RoboDK station: Celda_Soldadura_Estator_Grupo4_v05.rdk

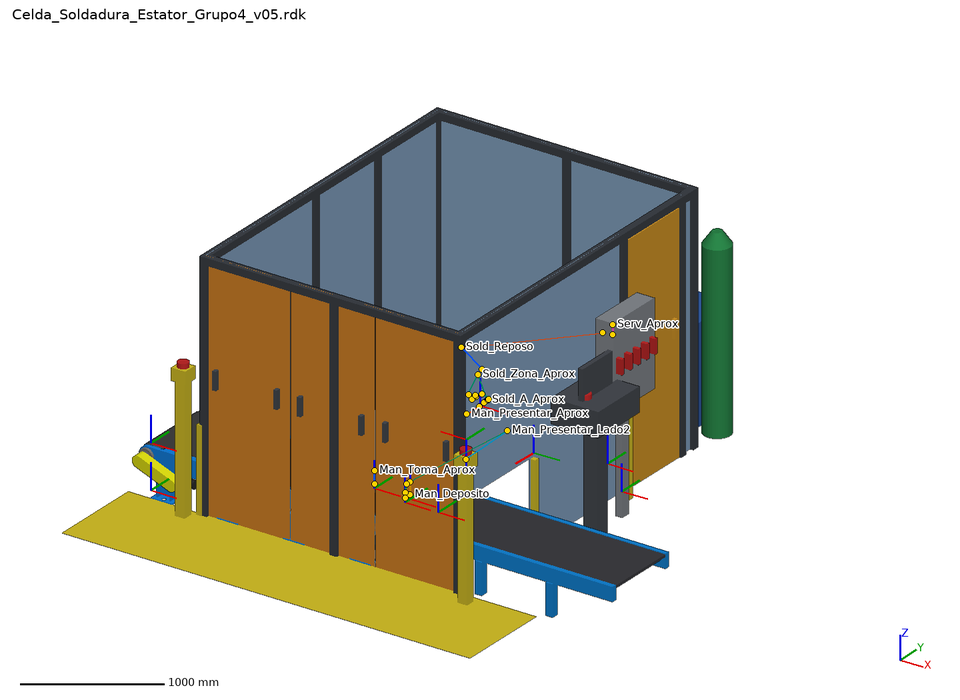
[picture v0: the station drawn from its stored meshes, robots at their saved joint values, targets as dots, program paths as lines]
Station Celda_Soldadura_Estator_Grupo4_v05 (saved by RoboDK 6.1.1). Poses are relative to the parent item; angles as X-Y-Z fixed-axis rotations.
Station parameters (name, value as stored): PIEZA_EN_TOMA, 0, PIEZA_PRESENTADA, 0, ARCO_TIG, 0, SOLDADURA_TERMINADA, 0, COORDINADOR_ACTIVO, 1, PERMISO_OPERACION, 0, ARRANQUE_ID, 0, ARRANQUE_ACK, 0, PARADA_ID, 0, PARADA_ACK, 0, AUTO_ACTIVO, 0, ESTADO_CONTROL, 0, CAUSA_RECHAZO, 0, PROXIMA_PIEZA, 1, PIEZA_ACTIVA, 0, CELDA_INICIALIZADA, 0, PIEZAS_COMPLETADAS, 0, LOTES_COMPLETADOS, 0, MODO_ID, 0, MODO_ACK, 0, MODO_SOLICITADO, 0, MODO_CONFIRMADO, 0, MODO_OBJETIVO, 0, MODO_EN_TRANSICION, 0, MODO_RESULTADO, 0, MODO_CAUSA, 0, MODO_ID_CAPTURADO, 0, MODO_CAPTURADO, 0, MODO_DESDE_AUTO, 0, MODO_ES_INTERVENCION, 0, MODO_CONOCIDO, 0, SENSORES_VALIDOS, 0, PIEZA_SUJETA_SENSOR, 0, IRB_EN_REPOSO, 0, CRB_EN_REPOSO, 0, IRB_EN_MANT, 0, CRB_EN_MANT, 0, CRB_EN_SERVICIO, 0, CINTA_DETENIDA, 0, IRB_DISPONIBLE, 0, CRB_DISPONIBLE, 0, CINTA_DISPONIBLE, 0, CONF_RESTITUCION, 0, FASE_PIEZA, 0, FASE_CAPTURADA, 0, PARO_CAUSA, 0, RECUP_PENDIENTE, 0, RECUPERAR_ID, 0, RECUPERAR_ACK, 0, PIEZAS_RETRABAJO, 0, RETRABAJO_ACTUAL, 0, SUJETA_CAPTURADA, 0, PIEZA_RESUELTA, 0, EMERGENCIA_SIM, 0, CORTINA_ENTRADA_SIM, 0, CORTINA_SALIDA_SIM, 0, PUERTA_ABIERTA_SIM, 0, OBJETIVO_PIEZAS, 0, PIEZAS_BUENAS, 0, PEDIDO_CUMPLIDO, 0, PEDIDOS_TERMINADOS, 0, REINICIAR_ID, 0, REINICIAR_ACK, 0, PEDIDO_PARADA, 0
  - frame Frame_Celda at (0, 0, 0) mm
    - frame Base_Manipulador_IRB1200 at (0, 0, 0) mm
      - robot ABB IRB 1200-7/0.7: 6 axes, payload 7 kg, reach 703 mm, repeatability 0.02 mm, weight 54 kg
          modified DH rows (alpha deg, a mm, theta deg, d mm): 0, 0, 0, 399; -90, 0, -90, 0; 0, 350, 0, 0; -90, 42, 0, 351; 90, 0, 0, 0; -90, 0, 180, 82
          joint limits [-170, -100, -200, -270, -130, -360] to [170, 135, 70, 270, 130, 360]; home [0, 0, 0, 0, 0, 0]; saved at [0, -20, 30, 0, 80, 0]
        - frame RobotiQ 2F-85 Gripper (Mechanism) Base at (0, 0, 0) mm
          - robot Pinza_2F85 (model RobotiQ 2F85): 1 axes, payload 5 kg
              joint limits [0] to [85]; home [85]; saved at [85]
        - tool TCP_Pinza, TCP at (0, 0, 150) mm
    - frame Base_Soldador_CRB1300 at (0, 1150, 0) mm, rotated rx 0 ry 0 rz -90 deg
      - robot ABB CRB 1300-10/1.15: 6 axes
          modified DH rows (alpha deg, a mm, theta deg, d mm): 0, 0, 0, 544; -90, 150, -90, 0; 0, 575, 0, 0; -90, 40, 0, 425; 90, 0, 0, 0; -90, 0, 180, 90
          joint limits [-180, -95, -210, -230, -130, -242] to [180, 155, 65, 230, 130, 242]; home [0, 0, 0, 0, 0, 0]; saved at [0, -10, 10, 0, 60, 0]
        - tool Antorcha_TIG, TCP at (0, 0, 207) mm, size 80 x 80 x 207 mm, geometry from antorcha_tig.stl
    - frame Base_Cinta_Pasante at (-1830, -860, 0) mm
      - robot Cinta_Pasante: 1 axes
          modified DH rows (alpha deg, a mm, theta deg, d mm): 0, 0, 0, 0 linear
          base shift (0, 0, 0) mm, rotated rx 0 ry 90 rz 0 deg
          joint limits [-900000] to [900000]; home [0]; saved at [0]
        - frame Frame_Banda at (0, 0, 0) mm
          - frame Frame_Piezas_Soldadas at (0, 0, 0) mm
          - object Estator_1 at (1680, 300, 0) mm, size 105 x 105 x 55 mm, geometry from paquete_estator.stl
          - object Estator_2 at (1380, 300, 0) mm, size 105 x 105 x 55 mm, geometry from paquete_estator.stl
          - object Estator_3 at (1080, 300, 0) mm, size 105 x 105 x 55 mm, geometry from paquete_estator.stl
          - object Estator_4 at (780, 300, 0) mm, size 105 x 105 x 55 mm, geometry from paquete_estator.stl
    - object Sensor_Pieza_En_Toma at (-150, -900, 396.5) mm, rotated rx 0 ry 0 rz 90 deg, size 683.3 x 45.2 x 12.5 mm, geometry from Laser-Sensor.stl
    - object Estacion_Servicio_Antorcha at (520, 1300, 0) mm, size 250 x 250 x 1000 mm, geometry from estacion_servicio_antorcha.stl
    - frame Frame_Cerramiento at (0, 0, 0) mm
      - frame Bisagra_Puerta at (850, 1000, 0) mm
        - object Puerta at (0, 0, 0) mm, size 60 x 700 x 1920 mm, geometry from puerta.stl
      - object Cerramiento_Estructura at (0, 0, 0) mm, size 2210 x 2870 x 2000 mm, geometry from cerramiento_estructura_v04.stl
      - object Cerramiento_Paneles at (0, 0, 0) mm, size 2154 x 2812 x 2000 mm, geometry from cerramiento_paneles_v04.stl
      - object Paneles_Desmontables_Sur at (0, 0, 0) mm, size 2140 x 4 x 2000 mm, geometry from paneles_desmontables_sur.stl
      - object Paneles_Desmontables_Manijas at (0, 0, 0) mm, size 1980 x 38 x 150 mm, geometry from paneles_desmontables_manijas.stl
      - object Cortina_Luz_Entrada at (-1330, 0, 0) mm, size 40 x 920 x 700 mm, geometry from cortina_luz_cinta_v04.stl
      - object Cortina_Luz_Salida at (880, 0, 0) mm, size 40 x 920 x 700 mm, geometry from cortina_luz_cinta_v04.stl
    - frame Frame_Soldadura at (0, 500, 620) mm
      - target Man_Presentar_Aprox (joint target) at (0, -157.5, 0) mm, rotated rx -90 ry 0 rz 0 deg; joints [90, -43.636, 55.703, 0, -12.068, -90] of ABB IRB 1200-7/0.7
      - target Man_Presentar_Lado1 (joint target) at (0, -7.5, 0) mm, rotated rx -90 ry 0 rz 0 deg; joints [90, -11.774, 38.724, 0, -26.95, -90] of ABB IRB 1200-7/0.7
      - target Man_Presentar_Lado2 (joint target) at (583, -500, 171) mm, rotated rx 0 ry 90 rz 0 deg; joints [90, -11.774, 38.724, 0, -26.95, 90] of ABB IRB 1200-7/0.7
      - target Man_Presentar_Aprox_Lado2 (joint target) at (583, -500, 171) mm, rotated rx 0 ry 90 rz 0 deg; joints [90, -43.636, 55.703, 0, -12.068, 90] of ABB IRB 1200-7/0.7
      - target Sold_Zona_Aprox (Cartesian target) at (0, -26.5, 250) mm, rotated rx 180 ry 0 rz 90 deg; joints [103.36, 41.617, 53.414, 0, -5.031, 103.36] of ABB CRB 1300-10/1.15
      - target Sold_A_Aprox (Cartesian target) at (78.2, -26.5, 78.2) mm, rotated rx -135 ry 0 rz 90 deg; joints [98.688, 74.302, 5.58, 7.491, 55.018, 91.856] of ABB CRB 1300-10/1.15
      - target Sold_A_Inicio (Cartesian target) at (49.91, -26.5, 49.91) mm, rotated rx -135 ry 0 rz 90 deg; joints [98.998, 76.411, 8.063, 8.245, 50.464, 91.119] of ABB CRB 1300-10/1.15
      - target Sold_A_Fin (Cartesian target) at (49.91, 26.5, 49.91) mm, rotated rx -135 ry 0 rz 90 deg; joints [102.751, 76.611, 6.557, 11.474, 51.681, 91.918] of ABB CRB 1300-10/1.15
      - target Sold_Transicion_Medio (Cartesian target) at (0, 26.5, 80) mm, rotated rx 180 ry 0 rz 90 deg; joints [108.748, 65.119, 46.933, 0, -22.052, 108.748] of ABB CRB 1300-10/1.15
      - target Sold_B_Inicio (Cartesian target) at (-49.91, 26.5, 49.91) mm, rotated rx 135 ry 0 rz 90 deg; joints [124.163, 102.688, 60.997, 205.222, 111.278, -54.665] of ABB CRB 1300-10/1.15
      - target Sold_B_Fin (Cartesian target) at (-49.91, -26.5, 49.91) mm, rotated rx 135 ry 0 rz 90 deg; joints [115.401, 107.202, 62.682, 200.569, 120.307, -60.716] of ABB CRB 1300-10/1.15
      - target Sold_B_Retiro (Cartesian target) at (-78.2, -26.5, 78.2) mm, rotated rx 135 ry 0 rz 90 deg; joints [-61.951, -75.264, -208.995, 23.114, 57.885, -82.141] of ABB CRB 1300-10/1.15
      - target Sold_A_Salida (Cartesian target) at (56.57, 26.5, 56.57) mm, rotated rx -135 ry 0 rz 90 deg; joints [102.647, 76.107, 6.003, 11.22, 52.72, 92.165] of ABB CRB 1300-10/1.15
      - target Sold_B_Entrada (Cartesian target) at (-56.57, 26.5, 56.57) mm, rotated rx 135 ry 0 rz 90 deg; joints [124.856, 103.181, 62.152, 205.935, 112.476, -53.248] of ABB CRB 1300-10/1.15
    - frame Frame_Toma_Cinta at (-150, -560, 366.5) mm
      - target Man_Toma_Aprox (joint target) at (0, 0, 135) mm, rotated rx 180 ry 0 rz 0 deg; joints [-104.995, 41.989, -47.307, 0, 95.319, 75.005] of ABB IRB 1200-7/0.7
      - target Man_Toma (joint target) at (0, 0, 35) mm, rotated rx 180 ry 0 rz 0 deg; joints [-104.995, 40.57, -28.656, 0, 78.086, 75.005] of ABB IRB 1200-7/0.7
    - frame Frame_Servicio at (520, 1300, 0) mm
      - target Serv_Aprox (Cartesian target) at (0, 60, 1050) mm, rotated rx 180 ry 0 rz 0 deg; joints [-125.65, 36.775, -52.607, 69.175, 38.577, -64.055] of ABB CRB 1300-10/1.15
      - target Serv_Verificacion_TCP (Cartesian target) at (0, 60, 973) mm, rotated rx 180 ry 0 rz 0 deg; joints [-125.65, 36.775, -52.607, 69.175, 38.577, -64.055] of ABB CRB 1300-10/1.15
      - target Serv_Cambio_Tungsteno (Cartesian target) at (0, -65, 1035) mm, rotated rx 180 ry 0 rz 0 deg; joints [-125.65, 36.775, -52.607, 69.175, 38.577, -64.055] of ABB CRB 1300-10/1.15
    - target Man_Reposo (joint target) at (583, 0, 791) mm, rotated rx 0 ry 90 rz 0 deg; joints [0, -20, 30, 0, 80, 0] of ABB IRB 1200-7/0.7
    - target Sold_Reposo (joint target) at (0, 278, 1159) mm, rotated rx 0 ry 90 rz -90 deg; joints [0, -10, 10, 0, 60, 0] of ABB CRB 1300-10/1.15
    - target Pinza_Abierta (joint target) at (536.92, 0, 791) mm, rotated rx 0 ry 90 rz 0 deg; joints [85] of Pinza_2F85
    - target Pinza_Cerrada (joint target) at (536.92, 0, 791) mm, rotated rx 0 ry 90 rz 0 deg; joints [0] of Pinza_2F85
    - target Pinza_Sujeta (joint target) at (536.92, 0, 791) mm, rotated rx 0 ry 90 rz 0 deg; joints [35] of Pinza_2F85
    - target Cinta_Posicion_1 (joint target) at (-1830, -860, 366.5) mm; joints [0] of Cinta_Pasante
    - target Cinta_Posicion_2 (joint target) at (-1830, -860, 366.5) mm; joints [300] of Cinta_Pasante
    - target Cinta_Posicion_3 (joint target) at (-1830, -860, 366.5) mm; joints [600] of Cinta_Pasante
    - target Cinta_Posicion_4 (joint target) at (-1830, -860, 366.5) mm; joints [900] of Cinta_Pasante
    - object Cinta_Salida_Banda at (0, 0, 0) mm, size 1880 x 600 x 20 mm, geometry from cinta_extension_banda.stl
    - object Cinta_Salida_Estructura at (0, 0, 0) mm, size 1880 x 700 x 371.5 mm, geometry from cinta_extension_estructura.stl
    - frame Frame_Deposito_Cinta at (150, -560, 366.5) mm
      - target Man_Deposito_Aprox (Cartesian target) at (0, 0, 135) mm, rotated rx 180 ry 0 rz 0 deg; joints [0, -20, 30, 0, 80, 0] of ABB IRB 1200-7/0.7
      - target Man_Deposito (Cartesian target) at (0, 0, 35) mm, rotated rx 180 ry 0 rz 0 deg; joints [0, -20, 30, 0, 80, 0] of ABB IRB 1200-7/0.7
    - target Cinta_Evacuacion (joint target) at (-1830, -860, 366.5) mm; joints [1750] of Cinta_Pasante
    - object Pasillo_Mantenimiento at (0, 0, 0) mm, size 3450 x 800 x 3 mm, geometry from pasillo_mantenimiento.stl
    - object Accionamiento_Cinta at (-1760, -80, 0) mm, size 140 x 320 x 296.5 mm, geometry from accionamiento_cinta.stl
    - object Accionamiento_Cinta_Resguardo at (-1760, -80, 0) mm, size 220 x 400 x 200 mm, geometry from accionamiento_cinta_resguardo.stl
    - object Tablero_LOTO at (1010, 700, 0) mm, size 150 x 500 x 1600 mm, geometry from tablero_loto.stl
    - object Tablero_LOTO_Seccionadores at (1010, 700, 0) mm, size 50 x 430 x 120 mm, geometry from tablero_loto_manijas.stl
    - object Panel_Operador at (1150, 250, 0) mm, size 400 x 500 x 1400 mm, geometry from panel_operador.stl
    - object Parada_Emergencia_Panel at (1150, 130, 0) mm, size 90 x 90 x 40 mm, geometry from parada_emergencia_hongo.stl
    - object Parada_Emergencia_Puerta_Poste at (930, 920, 0) mm, size 120 x 120 x 1150 mm, geometry from parada_emergencia_poste.stl
    - object Parada_Emergencia_Puerta at (930, 920, 0) mm, size 90 x 90 x 40 mm, geometry from parada_emergencia_hongo.stl
    - object Parada_Emergencia_Entrada_Poste at (-1420, -1060, 0) mm, size 120 x 120 x 1150 mm, geometry from parada_emergencia_poste.stl
    - object Parada_Emergencia_Entrada at (-1420, -1060, 0) mm, size 90 x 90 x 40 mm, geometry from parada_emergencia_hongo.stl
    - object Parada_Emergencia_Salida_Poste at (970, -1060, 0) mm, size 120 x 120 x 1150 mm, geometry from parada_emergencia_poste.stl
    - object Parada_Emergencia_Salida at (970, -1060, 0) mm, size 90 x 90 x 40 mm, geometry from parada_emergencia_hongo.stl
    - object Controlador_IRB1200 at (-800, 1950, 0) mm, size 600 x 500 x 1200 mm, geometry from gabinete_controlador.stl
    - object Controlador_CRB1300 at (-100, 1950, 0) mm, size 600 x 500 x 1200 mm, geometry from gabinete_controlador.stl
    - object Fuente_TIG at (500, 1950, 0) mm, size 400 x 600 x 800 mm, geometry from fuente_tig.stl
    - object Cilindro_Argon at (850, 2150, 0) mm, size 220 x 220 x 1550 mm, geometry from cilindro_argon.stl
    - target Man_Mantenimiento (joint target) at (233.25, 0, 476.3) mm, rotated rx 180 ry 0 rz -180 deg; joints [45, -30, 50, 0, 60, 0] of ABB IRB 1200-7/0.7
    - target Sold_Mantenimiento (joint target) at (0, 526.35, 893.05) mm, rotated rx 180 ry 30 rz 90 deg; joints [100, -30, 50, 0, 60, 0] of ABB CRB 1300-10/1.15
    - frame Frame_Deposito_Retrabajo at (150, -620, 366.5) mm
      - target Man_Retrabajo_Aprox (Cartesian target) at (0, 20, 135) mm, rotated rx 180 ry 0 rz 0 deg; joints [14.425, -18.655, 29.096, 0, 79.558, 14.425] of ABB IRB 1200-7/0.7
      - target Man_Retrabajo_Salida (Cartesian target) at (0, 0, 75) mm, rotated rx 180 ry 0 rz 0 deg; joints [14.425, -18.655, 29.096, 0, 79.558, 14.425] of ABB IRB 1200-7/0.7
      - target Man_Retrabajo (Cartesian target) at (0, 0, 35) mm, rotated rx 180 ry 0 rz 0 deg; joints [14.425, -18.655, 29.096, 0, 79.558, 14.425] of ABB IRB 1200-7/0.7
  - program Pinza_Abrir (2 instructions, listed below)
  - program Pinza_Cerrar (2 instructions, listed below)
  - program Pinza_Sujetar (2 instructions, listed below)
  - program Cinta_Avanzar_1 (4 instructions, listed below)
  - program Cinta_Avanzar_2 (4 instructions, listed below)
  - program Cinta_Avanzar_3 (4 instructions, listed below)
  - program Cinta_Avanzar_4 (4 instructions, listed below)
  - program Evento_Tomar_Pieza (2 instructions, listed below)
  - program Evento_Soltar_Pieza (2 instructions, listed below)
  - program Man_Ir_Reposo (4 instructions, listed below)
  - program Man_Tomar_Cinta (16 instructions, listed below)
  - program Man_Presentar_Lado1 (8 instructions, listed below)
  - program Man_Presentar_Lado2 (8 instructions, listed below)
  - program Sold_Ir_Reposo (4 instructions, listed below)
  - program Sold_Par_Cordones (38 instructions, listed below)
  - program Sold_Servicio_Antorcha (10 instructions, listed below)
  - program Inicio_Celda (8 instructions, listed below)
  - program Ciclo_Pieza_1 (15 instructions, listed below)
  - program Ciclo_Pieza_2 (15 instructions, listed below)
  - program Ciclo_Pieza_3 (15 instructions, listed below)
  - program Ciclo_Pieza_4 (17 instructions, listed below)
  - program Fin_Lote (6 instructions, listed below)
  - program Programa_Principal (8 instructions, listed below)
  - program Man_Depositar_Cinta (18 instructions, listed below)
  - program Cinta_Evacuar (2 instructions, listed below)
  - program Man_Ir_Mantenimiento (7 instructions, listed below)
  - program Sold_Ir_Mantenimiento (7 instructions, listed below)
  - program Preparar_Servicio_Antorcha (5 instructions, listed below)
  - program Parada_Entre_Piezas (7 instructions, listed below)
  - program Atender_Solicitud_Modo (598 instructions, listed below)
  - program Confirmar_Posicion_Modo (113 instructions, listed below)
  - program Man_Depositar_Retrabajo (19 instructions, listed below)
  - program Sold_Retirar (5 instructions, listed below)
  - program Recuperar_Desde_Lado1 (21 instructions, listed below)
  - program Recuperar_Desde_Lado2 (20 instructions, listed below)
  - program Recuperar_Deposito (18 instructions, listed below)
  - program Recuperar_Pieza (97 instructions, listed below)
  - program Cerrar_Pedido (14 instructions, listed below)
  - program Coordinador_Panel (275 instructions, listed below)
  - Python program Abrir_Panel_Operador (listed below)
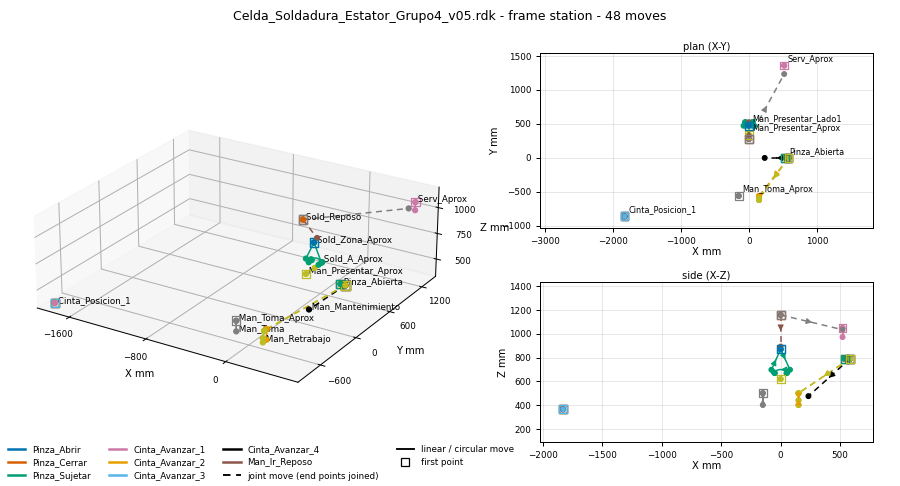
[picture p0: tool path of Celda_Soldadura_Estator_Grupo4_v05.rdk in frame station, 48 of 48 moves have a stored position in this frame; points joined in program order, loops and branches not executed]

--- program Pinza_Abrir (robot Pinza_2F85) ---
  Apertura máxima: reposo de la pinza
  MoveJ (Pinza_Abierta)

--- program Pinza_Cerrar (robot Pinza_2F85) ---
  Dedos juntos para entrar o salir del agujero del estator
  MoveJ (Pinza_Cerrada)

--- program Pinza_Sujetar (robot Pinza_2F85) ---
  Agarre interior: los dedos se abren contra el agujero de Ø55
  MoveJ (Pinza_Sujeta)

--- program Cinta_Avanzar_1 (robot Cinta_Pasante) ---
  Lleva el estator 1 del lote a la posición de toma
  MoveJ (Cinta_Posicion_1)
  Señal del sensor láser: hay pieza en la toma
  Set PIEZA_EN_TOMA=1

--- program Cinta_Avanzar_2 (robot Cinta_Pasante) ---
  Lleva el estator 2 del lote a la posición de toma
  MoveJ (Cinta_Posicion_2)
  Señal del sensor láser: hay pieza en la toma
  Set PIEZA_EN_TOMA=1

--- program Cinta_Avanzar_3 (robot Cinta_Pasante) ---
  Lleva el estator 3 del lote a la posición de toma
  MoveJ (Cinta_Posicion_3)
  Señal del sensor láser: hay pieza en la toma
  Set PIEZA_EN_TOMA=1

--- program Cinta_Avanzar_4 (robot Cinta_Pasante) ---
  Lleva el estator 4 del lote a la posición de toma
  MoveJ (Cinta_Posicion_4)
  Señal del sensor láser: hay pieza en la toma
  Set PIEZA_EN_TOMA=1

--- program Evento_Tomar_Pieza (robot ABB IRB 1200-7/0.7) ---
  Engancha a TCP_Pinza el estator que la pinza acaba de sujetar
  Adjuntar a TCP_Pinza

--- program Evento_Soltar_Pieza (robot ABB IRB 1200-7/0.7) ---
  Libera el estator sobre la banda (Frame_Piezas_Soldadas)
  Separar de TCP_Pinza

--- program Man_Ir_Reposo (robot ABB IRB 1200-7/0.7) ---
  Posición de reposo fuera de la zona de soldadura
  Est. herr: TCP_Pinza
  Establecer velocidad (1000.0 mm/s)
  MoveJ (Man_Reposo)

--- program Man_Tomar_Cinta (robot ABB IRB 1200-7/0.7) ---
  Toma el estator de la cinta con agarre interior
  Est. Ref.: Frame_Toma_Cinta
  Est. herr: TCP_Pinza
  Wait PIEZA_EN_TOMA=1
  Establecer velocidad (1000.0 mm/s)
  Suave(5)
  MoveJ (Man_Toma_Aprox)
  Llamar Pinza_Cerrar
  Suave(0)
  Establecer velocidad (100.0 mm/s)
  Entrada vertical en el agujero: MoveL para no rozar la pieza
  MoveL (Man_Toma)
  Llamar Pinza_Sujetar
  Llamar Evento_Tomar_Pieza
  Set PIEZA_EN_TOMA=0
  MoveL (Man_Toma_Aprox)

--- program Man_Presentar_Lado1 (robot ABB IRB 1200-7/0.7) ---
  Presenta las aristas A y B arriba, con el eje del estator hacia el soldador
  Est. Ref.: Frame_Soldadura
  Est. herr: TCP_Pinza
  Establecer velocidad (1000.0 mm/s)
  MoveJ (Man_Presentar_Aprox)
  Establecer velocidad (100.0 mm/s)
  MoveL (Man_Presentar_Lado1)
  Set PIEZA_PRESENTADA=1

--- program Man_Presentar_Lado2 (robot ABB IRB 1200-7/0.7) ---
  Gira 180° sobre el eje de la pinza (J6) para subir las aristas C y D
  Est. Ref.: Frame_Soldadura
  Est. herr: TCP_Pinza
  Wait SOLDADURA_TERMINADA=1
  Set SOLDADURA_TERMINADA=0
  Establecer velocidad (100.0 mm/s)
  MoveJ (Man_Presentar_Lado2)
  Set PIEZA_PRESENTADA=1

--- program Sold_Ir_Reposo (robot ABB CRB 1300-10/1.15) ---
  Reposo del soldador fuera del volumen de giro de la pieza
  Est. herr: Antorcha_TIG
  Establecer velocidad (1000.0 mm/s)
  MoveJ (Sold_Reposo)

--- program Sold_Par_Cordones (robot ABB CRB 1300-10/1.15) ---
  Suelda las dos aristas superiores del estator presentado
  Est. Ref.: Frame_Soldadura
  Est. herr: Antorcha_TIG
  Wait PIEZA_PRESENTADA=1
  Establecer velocidad (1000.0 mm/s)
  Suave(5)
  MoveJ (Sold_Zona_Aprox)
  Suave(0)
  Establecer velocidad (300.0 mm/s)
  Aproximación radial a la arista A
  MoveL (Sold_A_Aprox)
  Establecer velocidad (100.0 mm/s)
  MoveL (Sold_A_Inicio)
  Cordón A: arco encendido, avance recto a velocidad de soldadura
  Set ARCO_TIG=1
  Establecer velocidad (5.0 mm/s)
  MoveL (Sold_A_Fin)
  Set ARCO_TIG=0
  Establecer velocidad (100.0 mm/s)
  Separación radial: la punta sale del escalón antes de rodear la pieza
  MoveL (Sold_A_Salida)
  Establecer velocidad (200.0 mm/s)
  Transición en arco alrededor del eje del estator, a radio constante
  MoveC (Sold_Transicion_Medio, Sold_B_Entrada)
  Establecer velocidad (100.0 mm/s)
  MoveL (Sold_B_Inicio)
  Cordón B: avance recto en sentido contrario al A
  Set ARCO_TIG=1
  Establecer velocidad (5.0 mm/s)
  MoveL (Sold_B_Fin)
  Set ARCO_TIG=0
  Establecer velocidad (200.0 mm/s)
  MoveL (Sold_B_Retiro)
  Establecer velocidad (300.0 mm/s)
  MoveL (Sold_Zona_Aprox)
  Set PIEZA_PRESENTADA=0
  Set SOLDADURA_TERMINADA=1
  Llamar Sold_Ir_Reposo

--- program Sold_Servicio_Antorcha (robot ABB CRB 1300-10/1.15) ---
  Verificación del TCP al final de cada lote
  Est. Ref.: Frame_Servicio
  Est. herr: Antorcha_TIG
  Establecer velocidad (500.0 mm/s)
  MoveJ (Serv_Aprox)
  Establecer velocidad (100.0 mm/s)
  Bajada vertical hasta el cruce de los haces
  MoveL (Serv_Verificacion_TCP)
  MoveL (Serv_Aprox)
  Llamar Sold_Ir_Reposo

--- program Inicio_Celda (robot ABB IRB 1200-7/0.7) ---
  Estado inicial conocido: robots en reposo, pinza abierta, arco apagado
  Set ARCO_TIG=0
  Set PIEZA_EN_TOMA=0
  Set PIEZA_PRESENTADA=0
  Set SOLDADURA_TERMINADA=0
  Llamar Sold_Ir_Reposo
  Llamar Man_Ir_Reposo
  Llamar Pinza_Abrir

--- program Ciclo_Pieza_1 (robot ABB IRB 1200-7/0.7) ---
  Ciclo completo del estator 1: tomar, soldar 4 cordones, devolver a la banda
  Set FASE_PIEZA=1
  Llamar Cinta_Avanzar_1
  Set FASE_PIEZA=2
  Llamar Man_Tomar_Cinta
  Set FASE_PIEZA=3
  Llamar Man_Presentar_Lado1
  Set FASE_PIEZA=4
  Llamar Sold_Par_Cordones
  Set FASE_PIEZA=5
  Llamar Man_Presentar_Lado2
  Set FASE_PIEZA=6
  Llamar Sold_Par_Cordones
  Set FASE_PIEZA=7
  Llamar Man_Depositar_Cinta

--- program Ciclo_Pieza_2 (robot ABB IRB 1200-7/0.7) ---
  Ciclo completo del estator 2: tomar, soldar 4 cordones, devolver a la banda
  Set FASE_PIEZA=1
  Llamar Cinta_Avanzar_2
  Set FASE_PIEZA=2
  Llamar Man_Tomar_Cinta
  Set FASE_PIEZA=3
  Llamar Man_Presentar_Lado1
  Set FASE_PIEZA=4
  Llamar Sold_Par_Cordones
  Set FASE_PIEZA=5
  Llamar Man_Presentar_Lado2
  Set FASE_PIEZA=6
  Llamar Sold_Par_Cordones
  Set FASE_PIEZA=7
  Llamar Man_Depositar_Cinta

--- program Ciclo_Pieza_3 (robot ABB IRB 1200-7/0.7) ---
  Ciclo completo del estator 3: tomar, soldar 4 cordones, devolver a la banda
  Set FASE_PIEZA=1
  Llamar Cinta_Avanzar_3
  Set FASE_PIEZA=2
  Llamar Man_Tomar_Cinta
  Set FASE_PIEZA=3
  Llamar Man_Presentar_Lado1
  Set FASE_PIEZA=4
  Llamar Sold_Par_Cordones
  Set FASE_PIEZA=5
  Llamar Man_Presentar_Lado2
  Set FASE_PIEZA=6
  Llamar Sold_Par_Cordones
  Set FASE_PIEZA=7
  Llamar Man_Depositar_Cinta

--- program Ciclo_Pieza_4 (robot ABB IRB 1200-7/0.7) ---
  Ciclo completo del estator 4: tomar, soldar 4 cordones, devolver a la banda
  Set FASE_PIEZA=1
  Llamar Cinta_Avanzar_4
  Set FASE_PIEZA=2
  Llamar Man_Tomar_Cinta
  Set FASE_PIEZA=3
  Llamar Man_Presentar_Lado1
  Set FASE_PIEZA=4
  Llamar Sold_Par_Cordones
  Set FASE_PIEZA=5
  Llamar Man_Presentar_Lado2
  Set FASE_PIEZA=6
  Llamar Sold_Par_Cordones
  Set FASE_PIEZA=7
  Llamar Man_Depositar_Cinta
  Set FASE_PIEZA=8
  Llamar Man_Ir_Reposo

--- program Fin_Lote (robot ABB IRB 1200-7/0.7) ---
  Lote completo: verificación del TCP y evacuación de las piezas soldadas
  Llamar Sold_Servicio_Antorcha
  Llamar Cinta_Evacuar
  Reposición del lote (simula al operario que carga la entrada y retira la salida, afuera)
  Inicio Cinta_Pasante
  Mover objetos

--- program Programa_Principal (robot ABB IRB 1200-7/0.7) ---
  Celda de soldadura TIG de paquetes de estator - Grupo 4
  Ciclo nativo de un lote de 4 estatores; no necesita el panel
  Llamar Inicio_Celda
  Llamar Ciclo_Pieza_1
  Llamar Ciclo_Pieza_2
  Llamar Ciclo_Pieza_3
  Llamar Ciclo_Pieza_4
  Llamar Fin_Lote

--- program Man_Depositar_Cinta (robot ABB IRB 1200-7/0.7) ---
  Devuelve el estator soldado a la banda, aguas abajo de la toma
  Est. Ref.: Frame_Deposito_Cinta
  Est. herr: TCP_Pinza
  Wait SOLDADURA_TERMINADA=1
  Set SOLDADURA_TERMINADA=0
  Establecer velocidad (200.0 mm/s)
  MoveJ (Man_Presentar_Lado2)
  MoveL (Man_Presentar_Aprox_Lado2)
  Establecer velocidad (1000.0 mm/s)
  Suave(5)
  MoveJ (Man_Deposito_Aprox)
  Suave(0)
  Establecer velocidad (100.0 mm/s)
  Bajada vertical hasta apoyar la pieza en la banda
  MoveL (Man_Deposito)
  Llamar Pinza_Cerrar
  Llamar Evento_Soltar_Pieza
  MoveL (Man_Deposito_Aprox)

--- program Cinta_Evacuar (robot Cinta_Pasante) ---
  Avance final: saca el lote soldado por la salida de la celda
  MoveJ (Cinta_Evacuacion)

--- program Man_Ir_Mantenimiento (robot ABB IRB 1200-7/0.7) ---
  Lleva el IRB 1200 a su posición de mantenimiento: brazo plegado, herramienta hacia la puerta
  Se ejecuta en modo manual, con la celda detenida y nadie dentro
  Est. herr: TCP_Pinza
  Establecer velocidad (100.0 mm/s)
  MoveJ (Man_Reposo)
  MoveJ (Man_Mantenimiento)
  A continuación: bloqueo y etiquetado (LOTO) del IRB 1200, ver modos_y_mantenimiento.md §7

--- program Sold_Ir_Mantenimiento (robot ABB CRB 1300-10/1.15) ---
  Lleva el CRB 1300 a su posición de mantenimiento: brazo plegado, herramienta hacia la puerta
  Se ejecuta en modo manual, con la celda detenida y nadie dentro
  Est. herr: Antorcha_TIG
  Establecer velocidad (100.0 mm/s)
  MoveJ (Sold_Reposo)
  MoveJ (Sold_Mantenimiento)
  A continuación: bloqueo y etiquetado (LOTO) del CRB 1300, ver modos_y_mantenimiento.md §7

--- program Preparar_Servicio_Antorcha (robot ABB CRB 1300-10/1.15) ---
  Preparación sin pausa: acceso y aislamiento se tramitan después de posicionar
  Est. herr: Antorcha_TIG
  Establecer velocidad (100.0 mm/s)
  MoveJ (Sold_Reposo)
  MoveJ (Serv_Cambio_Tungsteno)

--- program Parada_Entre_Piezas (robot ABB IRB 1200-7/0.7) ---
  Set ARCO_TIG=0
  IF CRB_DISPONIBLE == 1
  Llamar Sold_Ir_Reposo
  END
  IF IRB_DISPONIBLE == 1
  Llamar Man_Ir_Reposo
  END

--- program Atender_Solicitud_Modo (robot ABB IRB 1200-7/0.7) ---
  IF MODO_ID != MODO_ACK
  MODO_ID_CAPTURADO = MODO_ID
  MODO_CAPTURADO = MODO_SOLICITADO
  Set MODO_RESULTADO=2
  Set MODO_CAUSA=0
  Set MODO_DESDE_AUTO=0
  Set MODO_ES_INTERVENCION=0
  Set MODO_CONOCIDO=0
  IF MODO_CAPTURADO == 0
  Set MODO_CONOCIDO=1
  END
  IF MODO_CAPTURADO == 1
  Set MODO_CONOCIDO=1
  END
  IF MODO_CAPTURADO == 1
  Set MODO_ES_INTERVENCION=1
  END
  IF MODO_CAPTURADO == 2
  Set MODO_CONOCIDO=1
  END
  IF MODO_CAPTURADO == 2
  Set MODO_ES_INTERVENCION=1
  END
  IF MODO_CAPTURADO == 3
  Set MODO_CONOCIDO=1
  END
  IF MODO_CAPTURADO == 3
  Set MODO_ES_INTERVENCION=1
  END
  IF MODO_CAPTURADO == 4
  Set MODO_CONOCIDO=1
  END
  IF MODO_CAPTURADO == 4
  Set MODO_ES_INTERVENCION=1
  END
  IF MODO_CAPTURADO == 5
  Set MODO_CONOCIDO=1
  END
  IF MODO_CAPTURADO == 5
  Set MODO_ES_INTERVENCION=1
  END
  IF MODO_CAPTURADO == 6
  Set MODO_CONOCIDO=1
  END
  IF MODO_CAPTURADO == 6
  Set MODO_ES_INTERVENCION=1
  END
  IF AUTO_ACTIVO == 1
  IF MODO_ES_INTERVENCION == 1
  Llamar Parada_Entre_Piezas
  Set AUTO_ACTIVO=0
  Set ESTADO_CONTROL=2
  Set MODO_DESDE_AUTO=1
  Set MODO_RESULTADO=3
  END
  END
  IF MODO_DESDE_AUTO == 0
  IF MODO_CONFIRMADO == 0
  IF MODO_CAPTURADO == 1
  IF IRB_DISPONIBLE == 0
  Set MODO_CAUSA=7
  END
  END
  END
  END
  IF MODO_DESDE_AUTO == 0
  IF MODO_CONFIRMADO == 0
  IF MODO_CAPTURADO == 2
  IF CRB_DISPONIBLE == 0
  Set MODO_CAUSA=7
  END
  END
  END
  END
  IF MODO_DESDE_AUTO == 0
  IF MODO_CONFIRMADO == 0
  IF MODO_CAPTURADO == 3
  IF IRB_DISPONIBLE == 0
  Set MODO_CAUSA=7
  END
  END
  END
  END
  IF MODO_DESDE_AUTO == 0
  IF MODO_CONFIRMADO == 0
  IF MODO_CAPTURADO == 3
  IF CRB_DISPONIBLE == 0
  Set MODO_CAUSA=7
  END
  END
  END
  END
  IF MODO_DESDE_AUTO == 0
  IF MODO_CONFIRMADO == 0
  IF MODO_CAPTURADO == 5
  IF CRB_DISPONIBLE == 0
  Set MODO_CAUSA=7
  END
  END
  END
  END
  IF MODO_DESDE_AUTO == 0
  IF MODO_ES_INTERVENCION == 1
  IF MODO_CONFIRMADO == 0
  IF MODO_CAPTURADO != 6
  IF IRB_EN_REPOSO == 0
  Set MODO_CAUSA=4
  END
  END
  END
  END
  END
  IF MODO_DESDE_AUTO == 0
  IF MODO_ES_INTERVENCION == 1
  IF MODO_CONFIRMADO == 0
  IF MODO_CAPTURADO != 6
  IF CRB_EN_REPOSO == 0
  Set MODO_CAUSA=4
  END
  END
  END
  END
  END
  IF MODO_DESDE_AUTO == 0
  IF MODO_ES_INTERVENCION == 1
  IF MODO_CONFIRMADO == 0
  IF MODO_CAPTURADO != 6
  IF PIEZA_SUJETA_SENSOR == 1
  Set MODO_CAUSA=5
  END
  END
  END
  END
  END
  IF MODO_DESDE_AUTO == 0
  IF MODO_ES_INTERVENCION == 1
  IF MODO_CONFIRMADO == 0
  IF MODO_CAPTURADO != 6
  IF PERMISO_OPERACION == 0
  Set MODO_CAUSA=1
  END
  END
  END
  END
  END
  IF MODO_DESDE_AUTO == 0
  IF MODO_CAPTURADO == 0
  IF MODO_CONFIRMADO == 1
  IF IRB_DISPONIBLE == 0
  Set MODO_CAUSA=7
  END
  END
  END
  END
  IF MODO_DESDE_AUTO == 0
  IF MODO_CAPTURADO == 0
  IF MODO_CONFIRMADO == 1
  IF IRB_EN_MANT == 0
  Set MODO_CAUSA=4
  END
  END
  END
  END
  IF MODO_DESDE_AUTO == 0
  IF MODO_CAPTURADO == 0
  IF MODO_CONFIRMADO == 1
  IF CRB_EN_REPOSO == 0
  Set MODO_CAUSA=4
  END
  END
  END
  END
  IF MODO_DESDE_AUTO == 0
  IF MODO_CAPTURADO == 0
  IF MODO_CONFIRMADO == 2
  IF CRB_DISPONIBLE == 0
  Set MODO_CAUSA=7
  END
  END
  END
  END
  IF MODO_DESDE_AUTO == 0
  IF MODO_CAPTURADO == 0
  IF MODO_CONFIRMADO == 2
  IF IRB_EN_REPOSO == 0
  Set MODO_CAUSA=4
  END
  END
  END
  END
  IF MODO_DESDE_AUTO == 0
  IF MODO_CAPTURADO == 0
  IF MODO_CONFIRMADO == 2
  IF CRB_EN_MANT == 0
  Set MODO_CAUSA=4
  END
  END
  END
  END
  IF MODO_DESDE_AUTO == 0
  IF MODO_CAPTURADO == 0
  IF MODO_CONFIRMADO == 3
  IF IRB_DISPONIBLE == 0
  Set MODO_CAUSA=7
  END
  END
  END
  END
  IF MODO_DESDE_AUTO == 0
  IF MODO_CAPTURADO == 0
  IF MODO_CONFIRMADO == 3
  IF CRB_DISPONIBLE == 0
  Set MODO_CAUSA=7
  END
  END
  END
  END
  IF MODO_DESDE_AUTO == 0
  IF MODO_CAPTURADO == 0
  IF MODO_CONFIRMADO == 3
  IF IRB_EN_MANT == 0
  Set MODO_CAUSA=4
  END
  END
  END
  END
  IF MODO_DESDE_AUTO == 0
  IF MODO_CAPTURADO == 0
  IF MODO_CONFIRMADO == 3
  IF CRB_EN_MANT == 0
  Set MODO_CAUSA=4
  END
  END
  END
  END
  IF MODO_DESDE_AUTO == 0
  IF MODO_CAPTURADO == 0
  IF MODO_CONFIRMADO == 4
  IF IRB_EN_REPOSO == 0
  Set MODO_CAUSA=4
  END
  END
  END
  END
  IF MODO_DESDE_AUTO == 0
  IF MODO_CAPTURADO == 0
  IF MODO_CONFIRMADO == 4
  IF CRB_EN_REPOSO == 0
  Set MODO_CAUSA=4
  END
  END
  END
  END
  IF MODO_DESDE_AUTO == 0
  IF MODO_CAPTURADO == 0
  IF MODO_CONFIRMADO == 5
  IF CRB_DISPONIBLE == 0
  Set MODO_CAUSA=7
  END
  END
  END
  END
  IF MODO_DESDE_AUTO == 0
  IF MODO_CAPTURADO == 0
  IF MODO_CONFIRMADO == 5
  IF IRB_EN_REPOSO == 0
  Set MODO_CAUSA=4
  END
  END
  END
  END
  IF MODO_DESDE_AUTO == 0
  IF MODO_CAPTURADO == 0
  IF MODO_CONFIRMADO == 5
  IF CRB_EN_SERVICIO == 0
  Set MODO_CAUSA=4
  END
  END
  END
  END
  IF MODO_DESDE_AUTO == 0
  IF MODO_CAPTURADO == 0
  IF MODO_CONFIRMADO == 6
  IF IRB_DISPONIBLE == 0
  Set MODO_CAUSA=7
  END
  END
  END
  END
  IF MODO_DESDE_AUTO == 0
  IF MODO_CAPTURADO == 0
  IF MODO_CONFIRMADO == 6
  IF CRB_DISPONIBLE == 0
  Set MODO_CAUSA=7
  END
  END
  END
  END
  IF MODO_DESDE_AUTO == 0
  IF MODO_CAPTURADO == 0
  IF MODO_CONFIRMADO == 6
  IF CINTA_DISPONIBLE == 0
  Set MODO_CAUSA=7
  END
  END
  END
  END
  IF MODO_DESDE_AUTO == 0
  IF MODO_CAPTURADO == 0
  IF MODO_CONFIRMADO == 6
  IF IRB_EN_REPOSO == 0
  Set MODO_CAUSA=4
  END
  END
  END
  END
  IF MODO_DESDE_AUTO == 0
  IF MODO_CAPTURADO == 0
  IF MODO_CONFIRMADO == 6
  IF CRB_EN_REPOSO == 0
  Set MODO_CAUSA=4
  END
  END
  END
  END
  IF MODO_DESDE_AUTO == 0
  IF MODO_CAPTURADO == 0
  IF MODO_CONFIRMADO != 0
  IF PIEZA_SUJETA_SENSOR == 1
  Set MODO_CAUSA=5
  END
  END
  END
  END
  IF MODO_DESDE_AUTO == 0
  IF MODO_CAPTURADO == 0
  IF MODO_CONFIRMADO != 0
  IF PERMISO_OPERACION == 0
  Set MODO_CAUSA=1
  END
  END
  END
  END
  IF MODO_DESDE_AUTO == 0
  IF MODO_CAPTURADO == 0
  IF MODO_CONFIRMADO != 0
  IF CONF_RESTITUCION == 0
  Set MODO_CAUSA=10
  END
  END
  END
  END
  IF MODO_DESDE_AUTO == 0
  IF MODO_CAPTURADO == 0
  IF MODO_CONFIRMADO == 0
  Set MODO_CAUSA=9
  END
  END
  END
  IF MODO_DESDE_AUTO == 0
  IF MODO_ES_INTERVENCION == 1
  IF MODO_CONFIRMADO != 0
  Set MODO_CAUSA=8
  END
  END
  END
  IF MODO_DESDE_AUTO == 0
  IF MODO_CONOCIDO == 1
  IF CINTA_DETENIDA == 0
  Set MODO_CAUSA=6
  END
  END
  END
  IF MODO_DESDE_AUTO == 0
  IF MODO_CONOCIDO == 1
  IF SENSORES_VALIDOS == 0
  Set MODO_CAUSA=3
  END
  END
  END
  IF MODO_DESDE_AUTO == 0
  IF MODO_CONOCIDO == 1
  IF MODO_EN_TRANSICION == 1
  Set MODO_CAUSA=2
  END
  END
  END
  IF MODO_DESDE_AUTO == 0
  IF MODO_CONOCIDO == 1
  IF RECUP_PENDIENTE == 1
  Set MODO_CAUSA=16
  END
  END
  END
  IF MODO_DESDE_AUTO == 0
  IF MODO_CONOCIDO == 1
  IF PARO_CAUSA != 0
  Set MODO_CAUSA=14
  END
  END
  END
  IF MODO_DESDE_AUTO == 0
  IF MODO_CONOCIDO == 0
  Set MODO_CAUSA=11
  END
  END
  IF MODO_DESDE_AUTO == 0
  IF MODO_CONOCIDO == 1
  IF MODO_CAUSA == 0
  IF MODO_CONFIRMADO == 0
  IF MODO_CAPTURADO == 1
  Set ARCO_TIG=0
  Set MODO_EN_TRANSICION=1
  Set ESTADO_CONTROL=4
  Llamar Man_Ir_Mantenimiento
  Set MODO_OBJETIVO=1
  Set MODO_RESULTADO=1
  END
  END
  END
  END
  END
  IF MODO_DESDE_AUTO == 0
  IF MODO_CONOCIDO == 1
  IF MODO_CAUSA == 0
  IF MODO_CONFIRMADO == 0
  IF MODO_CAPTURADO == 2
  Set ARCO_TIG=0
  Set MODO_EN_TRANSICION=1
  Set ESTADO_CONTROL=4
  Llamar Sold_Ir_Mantenimiento
  Set MODO_OBJETIVO=2
  Set MODO_RESULTADO=1
  END
  END
  END
  END
  END
  IF MODO_DESDE_AUTO == 0
  IF MODO_CONOCIDO == 1
  IF MODO_CAUSA == 0
  IF MODO_CONFIRMADO == 0
  IF MODO_CAPTURADO == 3
  Set ARCO_TIG=0
  Set MODO_EN_TRANSICION=1
  Set ESTADO_CONTROL=4
  Llamar Man_Ir_Mantenimiento
  Llamar Sold_Ir_Mantenimiento
  Set MODO_OBJETIVO=3
  Set MODO_RESULTADO=1
  END
  END
  END
  END
  END
  IF MODO_DESDE_AUTO == 0
  IF MODO_CONOCIDO == 1
  IF MODO_CAUSA == 0
  IF MODO_CONFIRMADO == 0
  IF MODO_CAPTURADO == 4
  Set ARCO_TIG=0
  Set MODO_EN_TRANSICION=1
  Set ESTADO_CONTROL=4
  Set MODO_OBJETIVO=4
  Set MODO_RESULTADO=1
  END
  END
  END
  END
  END
  IF MODO_DESDE_AUTO == 0
  IF MODO_CONOCIDO == 1
  IF MODO_CAUSA == 0
  IF MODO_CONFIRMADO == 0
  IF MODO_CAPTURADO == 5
  Set ARCO_TIG=0
  Set MODO_EN_TRANSICION=1
  Set ESTADO_CONTROL=4
  Llamar Preparar_Servicio_Antorcha
  Set MODO_OBJETIVO=5
  Set MODO_RESULTADO=1
  END
  END
  END
  END
  END
  IF MODO_DESDE_AUTO == 0
  IF MODO_CONOCIDO == 1
  IF MODO_CAUSA == 0
  IF MODO_CONFIRMADO == 0
  IF MODO_CAPTURADO == 6
  Set ARCO_TIG=0
  Set MODO_EN_TRANSICION=1
  Set ESTADO_CONTROL=4
  Set MODO_OBJETIVO=6
  Set MODO_RESULTADO=1
  END
  END
  END
  END
  END
  IF MODO_DESDE_AUTO == 0
  IF MODO_CONOCIDO == 1
  IF MODO_CAUSA == 0
  IF MODO_CAPTURADO == 0
  IF MODO_CONFIRMADO == 1
  Set MODO_EN_TRANSICION=1
  Set ESTADO_CONTROL=5
  Llamar Man_Ir_Reposo
  Set MODO_OBJETIVO=0
  Set MODO_RESULTADO=1
  Set CONF_RESTITUCION=0
  END
  END
  END
  END
  END
  IF MODO_DESDE_AUTO == 0
  IF MODO_CONOCIDO == 1
  IF MODO_CAUSA == 0
  IF MODO_CAPTURADO == 0
  IF MODO_CONFIRMADO == 2
  Set MODO_EN_TRANSICION=1
  Set ESTADO_CONTROL=5
  Llamar Sold_Ir_Reposo
  Set MODO_OBJETIVO=0
  Set MODO_RESULTADO=1
  Set CONF_RESTITUCION=0
  END
  END
  END
  END
  END
  IF MODO_DESDE_AUTO == 0
  IF MODO_CONOCIDO == 1
  IF MODO_CAUSA == 0
  IF MODO_CAPTURADO == 0
  IF MODO_CONFIRMADO == 3
  Set MODO_EN_TRANSICION=1
  Set ESTADO_CONTROL=5
  Llamar Sold_Ir_Reposo
  Llamar Man_Ir_Reposo
  Set MODO_OBJETIVO=0
  Set MODO_RESULTADO=1
  Set CONF_RESTITUCION=0
  END
  END
  END
  END
  END
  IF MODO_DESDE_AUTO == 0
  IF MODO_CONOCIDO == 1
  IF MODO_CAUSA == 0
  IF MODO_CAPTURADO == 0
  IF MODO_CONFIRMADO == 4
  Set MODO_EN_TRANSICION=1
  Set ESTADO_CONTROL=5
  Set MODO_OBJETIVO=0
  Set MODO_RESULTADO=1
  Set CONF_RESTITUCION=0
  END
  END
  END
  END
  END
  IF MODO_DESDE_AUTO == 0
  IF MODO_CONOCIDO == 1
  IF MODO_CAUSA == 0
  IF MODO_CAPTURADO == 0
  IF MODO_CONFIRMADO == 5
  Set MODO_EN_TRANSICION=1
  Set ESTADO_CONTROL=5
  Llamar Sold_Servicio_Antorcha
  Set MODO_OBJETIVO=0
  Set MODO_RESULTADO=1
  Set CONF_RESTITUCION=0
  END
  END
  END
  END
  END
  IF MODO_DESDE_AUTO == 0
  IF MODO_CONOCIDO == 1
  IF MODO_CAUSA == 0
  IF MODO_CAPTURADO == 0
  IF MODO_CONFIRMADO == 6
  Set MODO_EN_TRANSICION=1
  Set ESTADO_CONTROL=5
  Set MODO_OBJETIVO=0
  Set MODO_RESULTADO=1
  Set CONF_RESTITUCION=0
  END
  END
  END
  END
  END
  MODO_ACK = MODO_ID_CAPTURADO
  END

--- program Confirmar_Posicion_Modo (robot ABB IRB 1200-7/0.7) ---
  IF MODO_EN_TRANSICION == 1
  IF SENSORES_VALIDOS == 1
  IF CINTA_DETENIDA == 1
  IF PIEZA_SUJETA_SENSOR == 0
  IF MODO_OBJETIVO == 0
  IF IRB_EN_REPOSO == 1
  IF CRB_EN_REPOSO == 1
  Set MODO_CONFIRMADO=0
  Set MODO_EN_TRANSICION=0
  Set ESTADO_CONTROL=2
  END
  END
  END
  END
  END
  END
  END
  IF MODO_EN_TRANSICION == 1
  IF SENSORES_VALIDOS == 1
  IF CINTA_DETENIDA == 1
  IF PIEZA_SUJETA_SENSOR == 0
  IF MODO_OBJETIVO == 1
  IF IRB_EN_MANT == 1
  IF CRB_EN_REPOSO == 1
  Set MODO_CONFIRMADO=1
  Set MODO_EN_TRANSICION=0
  Set ESTADO_CONTROL=6
  END
  END
  END
  END
  END
  END
  END
  IF MODO_EN_TRANSICION == 1
  IF SENSORES_VALIDOS == 1
  IF CINTA_DETENIDA == 1
  IF PIEZA_SUJETA_SENSOR == 0
  IF MODO_OBJETIVO == 2
  IF IRB_EN_REPOSO == 1
  IF CRB_EN_MANT == 1
  Set MODO_CONFIRMADO=2
  Set MODO_EN_TRANSICION=0
  Set ESTADO_CONTROL=6
  END
  END
  END
  END
  END
  END
  END
  IF MODO_EN_TRANSICION == 1
  IF SENSORES_VALIDOS == 1
  IF CINTA_DETENIDA == 1
  IF PIEZA_SUJETA_SENSOR == 0
  IF MODO_OBJETIVO == 3
  IF IRB_EN_MANT == 1
  IF CRB_EN_MANT == 1
  Set MODO_CONFIRMADO=3
  Set MODO_EN_TRANSICION=0
  Set ESTADO_CONTROL=6
  END
  END
  END
  END
  END
  END
  END
  IF MODO_EN_TRANSICION == 1
  IF SENSORES_VALIDOS == 1
  IF CINTA_DETENIDA == 1
  IF PIEZA_SUJETA_SENSOR == 0
  IF MODO_OBJETIVO == 4
  IF IRB_EN_REPOSO == 1
  IF CRB_EN_REPOSO == 1
  Set MODO_CONFIRMADO=4
  Set MODO_EN_TRANSICION=0
  Set ESTADO_CONTROL=6
  END
  END
  END
  END
  END
  END
  END
  IF MODO_EN_TRANSICION == 1
  IF SENSORES_VALIDOS == 1
  IF CINTA_DETENIDA == 1
  IF PIEZA_SUJETA_SENSOR == 0
  IF MODO_OBJETIVO == 5
  IF IRB_EN_REPOSO == 1
  IF CRB_EN_SERVICIO == 1
  Set MODO_CONFIRMADO=5
  Set MODO_EN_TRANSICION=0
  Set ESTADO_CONTROL=6
  END
  END
  END
  END
  END
  END
  END
  IF MODO_EN_TRANSICION == 1
  IF SENSORES_VALIDOS == 1
  IF CINTA_DETENIDA == 1
  IF MODO_OBJETIVO == 6
  Set MODO_CONFIRMADO=6
  Set MODO_EN_TRANSICION=0
  Set ESTADO_CONTROL=6
  END
  END
  END
  END

--- program Man_Depositar_Retrabajo (robot ABB IRB 1200-7/0.7) ---
  Pieza de revisión o retrabajo: se deposita corrida hacia el borde derecho
  Est. Ref.: Frame_Deposito_Retrabajo
  Est. herr: TCP_Pinza
  Wait SOLDADURA_TERMINADA=1
  Set SOLDADURA_TERMINADA=0
  Establecer velocidad (200.0 mm/s)
  MoveJ (Man_Presentar_Lado2)
  MoveL (Man_Presentar_Aprox_Lado2)
  Establecer velocidad (1000.0 mm/s)
  Suave(5)
  MoveJ (Man_Retrabajo_Aprox)
  Suave(0)
  Establecer velocidad (100.0 mm/s)
  MoveL (Man_Retrabajo_Salida)
  MoveL (Man_Retrabajo)
  Llamar Pinza_Cerrar
  Llamar Evento_Soltar_Pieza
  MoveL (Man_Retrabajo_Salida)
  MoveL (Man_Retrabajo_Aprox)

--- program Sold_Retirar (robot ABB CRB 1300-10/1.15) ---
  Sale de la pieza en línea recta antes de ir a reposo
  Est. Ref.: Frame_Soldadura
  Est. herr: Antorcha_TIG
  Establecer velocidad (100.0 mm/s)
  MoveL (Sold_Zona_Aprox)

--- program Recuperar_Desde_Lado1 (robot ABB IRB 1200-7/0.7) ---
  Set ARCO_TIG=0
  Set PIEZA_PRESENTADA=0
  Set SOLDADURA_TERMINADA=0
  IF FASE_CAPTURADA == 4
  Llamar Sold_Retirar
  END
  IF FASE_CAPTURADA == 6
  Llamar Sold_Retirar
  END
  Llamar Sold_Ir_Reposo
  Llamar Man_Presentar_Lado1
  Llamar Sold_Par_Cordones
  Llamar Man_Presentar_Lado2
  Llamar Sold_Par_Cordones
  IF RETRABAJO_ACTUAL == 1
  Llamar Man_Depositar_Retrabajo
  END
  IF RETRABAJO_ACTUAL == 0
  Llamar Man_Depositar_Cinta
  END
  Llamar Man_Ir_Reposo

--- program Recuperar_Desde_Lado2 (robot ABB IRB 1200-7/0.7) ---
  Set ARCO_TIG=0
  Set PIEZA_PRESENTADA=0
  Set SOLDADURA_TERMINADA=0
  IF FASE_CAPTURADA == 4
  Llamar Sold_Retirar
  END
  IF FASE_CAPTURADA == 6
  Llamar Sold_Retirar
  END
  Llamar Sold_Ir_Reposo
  Set SOLDADURA_TERMINADA=1
  Llamar Man_Presentar_Lado2
  Llamar Sold_Par_Cordones
  IF RETRABAJO_ACTUAL == 1
  Llamar Man_Depositar_Retrabajo
  END
  IF RETRABAJO_ACTUAL == 0
  Llamar Man_Depositar_Cinta
  END
  Llamar Man_Ir_Reposo

--- program Recuperar_Deposito (robot ABB IRB 1200-7/0.7) ---
  Set ARCO_TIG=0
  Set PIEZA_PRESENTADA=0
  Set SOLDADURA_TERMINADA=0
  IF FASE_CAPTURADA == 4
  Llamar Sold_Retirar
  END
  IF FASE_CAPTURADA == 6
  Llamar Sold_Retirar
  END
  Llamar Sold_Ir_Reposo
  Set SOLDADURA_TERMINADA=1
  IF RETRABAJO_ACTUAL == 1
  Llamar Man_Depositar_Retrabajo
  END
  IF RETRABAJO_ACTUAL == 0
  Llamar Man_Depositar_Cinta
  END
  Llamar Man_Ir_Reposo

--- program Recuperar_Pieza (robot ABB IRB 1200-7/0.7) ---
  Retoma la pieza interrumpida; la soldadura se repite desde el par de cordones
  FASE_CAPTURADA = FASE_PIEZA
  Set RETRABAJO_ACTUAL=0
  Set PIEZA_RESUELTA=0
  Set SUJETA_CAPTURADA=0
  IF PIEZA_SUJETA_SENSOR == 1
  Set SUJETA_CAPTURADA=1
  END
  IF FASE_CAPTURADA == 4
  Set RETRABAJO_ACTUAL=1
  END
  IF FASE_CAPTURADA == 6
  Set RETRABAJO_ACTUAL=1
  END
  IF SUJETA_CAPTURADA == 0
  Set ARCO_TIG=0
  Set PIEZA_PRESENTADA=0
  Set SOLDADURA_TERMINADA=0
  IF FASE_CAPTURADA == 4
  Llamar Sold_Retirar
  END
  IF FASE_CAPTURADA == 6
  Llamar Sold_Retirar
  END
  Llamar Sold_Ir_Reposo
  Llamar Man_Ir_Reposo
  Llamar Pinza_Abrir
  IF FASE_CAPTURADA == 7
  Set PIEZA_RESUELTA=1
  END
  IF FASE_CAPTURADA == 8
  Set PIEZA_RESUELTA=1
  END
  END
  IF SUJETA_CAPTURADA == 1
  IF FASE_CAPTURADA == 1
  Llamar Recuperar_Desde_Lado1
  Set PIEZA_RESUELTA=1
  END
  END
  IF SUJETA_CAPTURADA == 1
  IF FASE_CAPTURADA == 2
  Llamar Recuperar_Desde_Lado1
  Set PIEZA_RESUELTA=1
  END
  END
  IF SUJETA_CAPTURADA == 1
  IF FASE_CAPTURADA == 3
  Llamar Recuperar_Desde_Lado1
  Set PIEZA_RESUELTA=1
  END
  END
  IF SUJETA_CAPTURADA == 1
  IF FASE_CAPTURADA == 4
  Llamar Recuperar_Desde_Lado1
  Set PIEZA_RESUELTA=1
  END
  END
  IF SUJETA_CAPTURADA == 1
  IF FASE_CAPTURADA == 5
  Llamar Recuperar_Desde_Lado2
  Set PIEZA_RESUELTA=1
  END
  END
  IF SUJETA_CAPTURADA == 1
  IF FASE_CAPTURADA == 6
  Llamar Recuperar_Desde_Lado2
  Set PIEZA_RESUELTA=1
  END
  END
  IF SUJETA_CAPTURADA == 1
  IF FASE_CAPTURADA == 7
  Llamar Recuperar_Deposito
  Set PIEZA_RESUELTA=1
  END
  END
  IF SUJETA_CAPTURADA == 1
  IF FASE_CAPTURADA == 8
  Llamar Recuperar_Deposito
  Set PIEZA_RESUELTA=1
  END
  END
  IF PIEZA_RESUELTA == 1
  IF PIEZA_ACTIVA != 0
  PROXIMA_PIEZA = PROXIMA_PIEZA + 1
  PIEZAS_COMPLETADAS = PIEZAS_COMPLETADAS + 1
  END
  END
  IF RETRABAJO_ACTUAL == 1
  IF PIEZA_RESUELTA == 1
  PIEZAS_RETRABAJO = PIEZAS_RETRABAJO + 1
  END
  END
  Set PIEZA_ACTIVA=0
  Set FASE_PIEZA=0
  Set MODO_EN_TRANSICION=0
  Set MODO_OBJETIVO=0

--- program Cerrar_Pedido (robot ABB IRB 1200-7/0.7) ---
  Evacúa y repone las piezas, aunque el lote esté incompleto, y deja todo en cero
  IF PROXIMA_PIEZA != 1
  Llamar Man_Ir_Reposo
  Llamar Fin_Lote
  END
  Set PIEZAS_COMPLETADAS=0
  Set PIEZAS_RETRABAJO=0
  Set PIEZAS_BUENAS=0
  Set LOTES_COMPLETADOS=0
  Set AUTO_ACTIVO=0
  Set PEDIDO_CUMPLIDO=0
  Set PROXIMA_PIEZA=1
  Set ESTADO_CONTROL=9
  PEDIDOS_TERMINADOS = PEDIDOS_TERMINADOS + 1

--- program Coordinador_Panel (robot ABB IRB 1200-7/0.7) ---
  Coordinador v05: iniciar desde RoboDK; mandos por señales. PERMISO_OPERACION no es una parada inmediata de protección.
  IF AUTO_ACTIVO == 1
  Set RECUP_PENDIENTE=1
  Set AUTO_ACTIVO=0
  Set ESTADO_CONTROL=7
  END
  IF PIEZA_ACTIVA != 0
  Set RECUP_PENDIENTE=1
  Set AUTO_ACTIVO=0
  Set ESTADO_CONTROL=7
  END
  IF MODO_EN_TRANSICION == 1
  Set RECUP_PENDIENTE=1
  Set AUTO_ACTIVO=0
  Set ESTADO_CONTROL=7
  END
  WHILE COORDINADOR_ACTIVO == 1
  Set PEDIDO_PARADA=0
  IF PARADA_ID != PARADA_ACK
  Set PEDIDO_PARADA=1
  END
  IF PEDIDO_PARADA == 1
  IF ARRANQUE_ID != ARRANQUE_ACK
  Set CAUSA_RECHAZO=13
  ARRANQUE_ACK = ARRANQUE_ID
  END
  IF AUTO_ACTIVO == 1
  Llamar Parada_Entre_Piezas
  END
  Set AUTO_ACTIVO=0
  Set ESTADO_CONTROL=2
  PARADA_ACK = PARADA_ID
  END
  Llamar Atender_Solicitud_Modo
  Llamar Confirmar_Posicion_Modo
  IF PEDIDO_PARADA == 0
  IF ARRANQUE_ID != ARRANQUE_ACK
  Set CAUSA_RECHAZO=0
  IF CINTA_DISPONIBLE == 0
  Set CAUSA_RECHAZO=7
  END
  IF CRB_DISPONIBLE == 0
  Set CAUSA_RECHAZO=7
  END
  IF IRB_DISPONIBLE == 0
  Set CAUSA_RECHAZO=7
  END
  IF CINTA_DETENIDA == 0
  Set CAUSA_RECHAZO=6
  END
  IF PIEZA_SUJETA_SENSOR == 1
  Set CAUSA_RECHAZO=5
  END
  IF CRB_EN_REPOSO == 0
  Set CAUSA_RECHAZO=4
  END
  IF IRB_EN_REPOSO == 0
  Set CAUSA_RECHAZO=4
  END
  IF SENSORES_VALIDOS == 0
  Set CAUSA_RECHAZO=3
  END
  IF MODO_CONFIRMADO != 0
  Set CAUSA_RECHAZO=8
  END
  IF MODO_EN_TRANSICION == 1
  Set CAUSA_RECHAZO=2
  END
  IF PERMISO_OPERACION == 0
  Set CAUSA_RECHAZO=1
  END
  IF AUTO_ACTIVO == 1
  Set CAUSA_RECHAZO=12
  END
  IF RECUP_PENDIENTE == 1
  Set CAUSA_RECHAZO=16
  END
  IF CORTINA_ENTRADA_SIM == 1
  Set CAUSA_RECHAZO=15
  END
  IF CORTINA_SALIDA_SIM == 1
  Set CAUSA_RECHAZO=15
  END
  IF PUERTA_ABIERTA_SIM == 1
  Set CAUSA_RECHAZO=15
  END
  IF PARO_CAUSA != 0
  Set CAUSA_RECHAZO=14
  END
  ARRANQUE_ACK = ARRANQUE_ID
  IF CAUSA_RECHAZO == 0
  IF CELDA_INICIALIZADA == 0
  Llamar Inicio_Celda
  Set CELDA_INICIALIZADA=1
  END
  Set AUTO_ACTIVO=1
  Set ESTADO_CONTROL=1
  END
  END
  END
  IF RECUPERAR_ID != RECUPERAR_ACK
  Set CAUSA_RECHAZO=0
  IF CRB_DISPONIBLE == 0
  Set CAUSA_RECHAZO=7
  END
  IF IRB_DISPONIBLE == 0
  Set CAUSA_RECHAZO=7
  END
  IF SENSORES_VALIDOS == 0
  Set CAUSA_RECHAZO=3
  END
  IF PERMISO_OPERACION == 0
  Set CAUSA_RECHAZO=1
  END
  IF RECUP_PENDIENTE == 0
  Set CAUSA_RECHAZO=17
  END
  IF CORTINA_ENTRADA_SIM == 1
  Set CAUSA_RECHAZO=15
  END
  IF CORTINA_SALIDA_SIM == 1
  Set CAUSA_RECHAZO=15
  END
  IF PUERTA_ABIERTA_SIM == 1
  Set CAUSA_RECHAZO=15
  END
  IF PARO_CAUSA != 0
  Set CAUSA_RECHAZO=14
  END
  RECUPERAR_ACK = RECUPERAR_ID
  IF CAUSA_RECHAZO == 0
  Set ESTADO_CONTROL=8
  Llamar Recuperar_Pieza
  Set RECUP_PENDIENTE=0
  Set ESTADO_CONTROL=2
  END
  END
  IF AUTO_ACTIVO == 1
  IF PERMISO_OPERACION == 0
  Llamar Parada_Entre_Piezas
  Set AUTO_ACTIVO=0
  Set ESTADO_CONTROL=3
  END
  END
  IF AUTO_ACTIVO == 1
  IF SENSORES_VALIDOS == 0
  Llamar Parada_Entre_Piezas
  Set AUTO_ACTIVO=0
  Set ESTADO_CONTROL=3
  END
  END
  IF AUTO_ACTIVO == 1
  IF IRB_DISPONIBLE == 0
  Llamar Parada_Entre_Piezas
  Set AUTO_ACTIVO=0
  Set ESTADO_CONTROL=3
  END
  END
  IF AUTO_ACTIVO == 1
  IF CRB_DISPONIBLE == 0
  Llamar Parada_Entre_Piezas
  Set AUTO_ACTIVO=0
  Set ESTADO_CONTROL=3
  END
  END
  IF AUTO_ACTIVO == 1
  IF CINTA_DISPONIBLE == 0
  Llamar Parada_Entre_Piezas
  Set AUTO_ACTIVO=0
  Set ESTADO_CONTROL=3
  END
  END
  PIEZAS_BUENAS = PIEZAS_COMPLETADAS - PIEZAS_RETRABAJO
  IF AUTO_ACTIVO == 1
  IF OBJETIVO_PIEZAS > 0
  IF PIEZAS_BUENAS >= OBJETIVO_PIEZAS
  Set PEDIDO_CUMPLIDO=1
  END
  END
  END
  IF REINICIAR_ID != REINICIAR_ACK
  Set CAUSA_RECHAZO=0
  IF CINTA_DISPONIBLE == 0
  Set CAUSA_RECHAZO=7
  END
  IF CINTA_DETENIDA == 0
  Set CAUSA_RECHAZO=6
  END
  IF PIEZA_SUJETA_SENSOR == 1
  Set CAUSA_RECHAZO=5
  END
  IF CRB_EN_REPOSO == 0
  Set CAUSA_RECHAZO=4
  END
  IF IRB_EN_REPOSO == 0
  Set CAUSA_RECHAZO=4
  END
  IF SENSORES_VALIDOS == 0
  Set CAUSA_RECHAZO=3
  END
  IF MODO_CONFIRMADO != 0
  Set CAUSA_RECHAZO=8
  END
  IF PERMISO_OPERACION == 0
  Set CAUSA_RECHAZO=1
  END
  IF AUTO_ACTIVO == 1
  Set CAUSA_RECHAZO=12
  END
  IF RECUP_PENDIENTE == 1
  Set CAUSA_RECHAZO=16
  END
  IF CORTINA_ENTRADA_SIM == 1
  Set CAUSA_RECHAZO=15
  END
  IF CORTINA_SALIDA_SIM == 1
  Set CAUSA_RECHAZO=15
  END
  IF PUERTA_ABIERTA_SIM == 1
  Set CAUSA_RECHAZO=15
  END
  IF PARO_CAUSA != 0
  Set CAUSA_RECHAZO=14
  END
  REINICIAR_ACK = REINICIAR_ID
  IF CAUSA_RECHAZO == 0
  Set PEDIDO_CUMPLIDO=1
  END
  END
  IF PEDIDO_CUMPLIDO == 1
  IF PARO_CAUSA == 0
  IF RECUP_PENDIENTE == 0
  Llamar Cerrar_Pedido
  END
  END
  END
  IF AUTO_ACTIVO == 1
  INDICE_CAPTURADO = PROXIMA_PIEZA
  IF INDICE_CAPTURADO == 1
  Set PIEZA_ACTIVA=1
  Llamar Ciclo_Pieza_1
  Set PIEZA_ACTIVA=0
  Set PROXIMA_PIEZA=2
  PIEZAS_COMPLETADAS = PIEZAS_COMPLETADAS + 1
  END
  IF INDICE_CAPTURADO == 2
  Set PIEZA_ACTIVA=2
  Llamar Ciclo_Pieza_2
  Set PIEZA_ACTIVA=0
  Set PROXIMA_PIEZA=3
  PIEZAS_COMPLETADAS = PIEZAS_COMPLETADAS + 1
  END
  IF INDICE_CAPTURADO == 3
  Set PIEZA_ACTIVA=3
  Llamar Ciclo_Pieza_3
  Set PIEZA_ACTIVA=0
  Set PROXIMA_PIEZA=4
  PIEZAS_COMPLETADAS = PIEZAS_COMPLETADAS + 1
  END
  IF INDICE_CAPTURADO == 4
  Set PIEZA_ACTIVA=4
  Llamar Ciclo_Pieza_4
  Set PIEZA_ACTIVA=0
  Set PROXIMA_PIEZA=5
  PIEZAS_COMPLETADAS = PIEZAS_COMPLETADAS + 1
  END
  IF INDICE_CAPTURADO == 5
  Llamar Fin_Lote
  LOTES_COMPLETADOS = LOTES_COMPLETADOS + 1
  Set PROXIMA_PIEZA=1
  END
  END
  Pausa 100 ms
  END
  Set AUTO_ACTIVO=0

--- Python program Abrir_Panel_Operador ---
"""Panel de operador de la celda. Generado por empaquetar_panel.py: no editar aquí.

Se ejecuta con doble clic en RoboDK. Solo lee y escribe señales: no mueve robots ni la cinta.
"""
import os
import subprocess
import sys

# RoboDK puede tener configurado otro Python; PySide2 viene con el que trae la instalación.
PYTHON_ROBODK = r"C:\RoboDK\Python-Embedded\python.exe"
try:
    import PySide2
except ImportError:
    if os.path.exists(PYTHON_ROBODK) and os.path.normcase(sys.executable) != os.path.normcase(PYTHON_ROBODK):
        sys.exit(subprocess.call([PYTHON_ROBODK, __file__]))
    from robodk.robolink import Robolink
    Robolink().ShowMessage("El panel necesita PySide2, incluido en el Python de RoboDK 6.1.1.")
    sys.exit(1)

from enum import Enum
from dataclasses import dataclass
import hashlib
import hmac
import os
from pathlib import Path
import sqlite3
import time
import argparse
import math
import sys
from robodk.robolink import Robolink, ITEM_TYPE_ROBOT, ITEM_TYPE_TOOL, ITEM_TYPE_TARGET
import queue
import socket
from PySide2.QtCore import QThread, Signal
from robodk.robolink import Robolink, ITEM_TYPE_PROGRAM, ITEM_TYPE_ROBOT
from PySide2.QtCore import QPointF, QRectF, Qt, Signal
from PySide2.QtGui import QBrush, QColor, QFont, QPainter, QPen
from PySide2.QtWidgets import QSizePolicy, QWidget
from datetime import datetime
from PySide2.QtCore import QEvent, Qt, QTimer
from PySide2.QtWidgets import (QAbstractItemView, QCheckBox, QComboBox, QDialog, QFormLayout, QFrame,
                               QGridLayout, QGroupBox, QHBoxLayout, QHeaderView, QInputDialog,
                               QLabel, QLineEdit, QMainWindow, QMessageBox, QPushButton,
                               QSpinBox, QStackedWidget, QTableWidget, QTableWidgetItem, QTabWidget,
                               QTextBrowser, QVBoxLayout, QWidget)
from PySide2.QtWidgets import QApplication

CAUSAS = {
    0: "Sin causa de rechazo",
    1: "Sin permiso de operación",
    2: "Cambio de modo en curso",
    3: "Sensores no válidos",
    4: "Equipo fuera de la posición requerida",
    5: "Pieza sujeta",
    6: "Cinta en movimiento",
    7: "Equipo no disponible",
    8: "Hay un modo activo",
    9: "No hay modo del cual regresar",
    10: "Falta confirmar la restitución",
    11: "Modo desconocido",
    12: "Producción activa",
    13: "Arranque simultáneo con una parada",
    14: "Parada activa sin rearmar",
    15: "Resguardo abierto",
    16: "Recuperación pendiente",
    17: "No hay nada que recuperar",
}

# --- permisos.py ---

PRODUCCION = "produccion"

MANTENIMIENTO = "mantenimiento"

ADMINISTRADOR = "administrador"

PERFILES = (PRODUCCION, MANTENIMIENTO, ADMINISTRADOR)

class Op(Enum):
    ARRANQUE = "Arranque"
    PARADA = "Parada normal"
    PREPARAR_MODO = "Preparar modo"
    REGRESAR_MODO = "Regresar a producción"
    ENTRADA_SIMULADA = "Entrada simulada"
    ADMINISTRAR = "Administrar cuentas"
    EMERGENCIA = "Pulsador de emergencia"
    RESGUARDO = "Cortina o puerta"
    REARME = "Rearme"
    RECUPERAR = "Recuperación"
    REINICIAR = "Reinicio de lote"
    OBJETIVO = "Objetivo de piezas"

MATRIZ = {
    PRODUCCION: {Op.ARRANQUE, Op.PARADA, Op.EMERGENCIA, Op.RESGUARDO, Op.REARME, Op.OBJETIVO},
    MANTENIMIENTO: {Op.PARADA, Op.PREPARAR_MODO, Op.REGRESAR_MODO, Op.ENTRADA_SIMULADA, Op.EMERGENCIA,
                    Op.RESGUARDO, Op.REARME, Op.RECUPERAR, Op.REINICIAR},
    ADMINISTRADOR: {Op.PARADA, Op.ADMINISTRAR, Op.EMERGENCIA, Op.RESGUARDO},
}

MODOS = {
    1: "IRB 1200 y pinza",
    2: "CRB 1300",
    3: "Ambos robots",
    4: "Cinta",
    5: "Servicio de antorcha",
    6: "Correctivo sin movimiento",
}

TIPOS_INTERVENCION = ("Preventivo", "Correctivo")

ENTRADAS_SIMULADAS = ("PERMISO_OPERACION", "IRB_DISPONIBLE", "CRB_DISPONIBLE", "CINTA_DISPONIBLE")

RESGUARDOS = {"CORTINA_ENTRADA_SIM": 2, "CORTINA_SALIDA_SIM": 2, "PUERTA_ABIERTA_SIM": 3}

CAUSAS_PARO = {1: "Emergencia", 2: "Cortina de luz", 3: "Puerta abierta"}

OBJETIVO_MAXIMO = 9999

def permitido(perfil, operacion):
    return operacion in MATRIZ.get(perfil, ())

# --- cuentas.py ---

INACTIVIDAD_S = 15 * 60

INTENTOS_MAXIMOS = 5

BLOQUEO_S = 5 * 60

CLAVE_MINIMA = 8

SCRYPT_N, SCRYPT_R, SCRYPT_P = 2 ** 15, 8, 3

CUENTAS_INICIALES = (
    ("admin", "Administrador", ADMINISTRADOR, "admin"),
    ("mantenimiento", "Mantenimiento", MANTENIMIENTO, "mantenimiento"),
    ("produccion", "Producción", PRODUCCION, "produccion"),
)

FALLO_ACCESO = "Usuario o contraseña incorrectos, o acceso bloqueado temporalmente."

def ruta_datos():
    """La estación se entrega sola: la base se crea en los datos de quien usa el panel."""
    base = Path(os.environ.get("LOCALAPPDATA") or Path.home()) / "Celda_Soldadura_Grupo4"
    base.mkdir(parents=True, exist_ok=True)
    return base / "panel.db"

class ErrorCuenta(Exception):
    pass

@dataclass
class Sesion:
    usuario: str
    nombre: str
    perfil: str
    ultima_actividad: float
    clave_por_defecto: bool
    cerrada: bool = False

def _derivar(clave, sal, n, r, p):
    return hashlib.scrypt(clave.encode("utf-8"), salt=sal, n=n, r=r, p=p,
                          maxmem=128 * r * n * 2, dklen=32)

def generar_hash(clave):
    sal = os.urandom(16)
    derivada = _derivar(clave, sal, SCRYPT_N, SCRYPT_R, SCRYPT_P)
    return f"scrypt${SCRYPT_N}${SCRYPT_R}${SCRYPT_P}${sal.hex()}${derivada.hex()}"

def comprobar_hash(clave, guardado):
    _, n, r, p, sal, derivada = guardado.split("$")
    calculada = _derivar(clave, bytes.fromhex(sal), int(n), int(r), int(p))
    return hmac.compare_digest(calculada, bytes.fromhex(derivada))

class Cuentas:
    def __init__(self, ruta, reloj=time.time):
        self.reloj = reloj
        self.db = sqlite3.connect(str(ruta))
        self.db.row_factory = sqlite3.Row
        self.db.executescript("""
            CREATE TABLE IF NOT EXISTS usuarios (
                usuario TEXT PRIMARY KEY, nombre TEXT NOT NULL, perfil TEXT NOT NULL,
                clave TEXT NOT NULL, activo INTEGER NOT NULL DEFAULT 1,
                clave_por_defecto INTEGER NOT NULL DEFAULT 0,
                intentos INTEGER NOT NULL DEFAULT 0, bloqueado_hasta REAL NOT NULL DEFAULT 0,
                creado REAL NOT NULL);
            CREATE TABLE IF NOT EXISTS registro (
                id INTEGER PRIMARY KEY AUTOINCREMENT, fecha REAL NOT NULL, usuario TEXT NOT NULL,
                perfil TEXT NOT NULL, operacion TEXT NOT NULL, detalle TEXT NOT NULL,
                resultado TEXT NOT NULL);
        """)
        if not self.db.execute("SELECT 1 FROM usuarios LIMIT 1").fetchone():
            for usuario, nombre, perfil, clave in CUENTAS_INICIALES:
                self._insertar(usuario, nombre, perfil, clave, por_defecto=1)
            self.registrar("sistema", "-", "Crear base", "Cuentas iniciales", "Hecho")
        self._hash_ficticio = generar_hash(os.urandom(8).hex())

    def _insertar(self, usuario, nombre, perfil, clave, por_defecto=0):
        self.db.execute("INSERT INTO usuarios (usuario, nombre, perfil, clave, clave_por_defecto, "
                        "creado) VALUES (?, ?, ?, ?, ?, ?)",
                        (usuario, nombre, perfil, generar_hash(clave), por_defecto, self.reloj()))
        self.db.commit()

    def _fila(self, usuario):
        return self.db.execute("SELECT * FROM usuarios WHERE usuario = ?", (usuario,)).fetchone()

    def registrar(self, usuario, perfil, operacion, detalle, resultado):
        self.db.execute("INSERT INTO registro (fecha, usuario, perfil, operacion, detalle, resultado)"
                        " VALUES (?, ?, ?, ?, ?, ?)",
                        (self.reloj(), usuario, perfil, operacion, detalle, resultado))
        self.db.commit()

    def leer_registro(self, limite=200):
        return self.db.execute("SELECT * FROM registro ORDER BY id DESC LIMIT ?", (limite,)).fetchall()

    def autenticar(self, usuario, clave):
        """Devuelve una Sesion o None; el motivo del fallo no se revela a quien intenta entrar."""
        fila = self._fila(usuario)
        ahora = self.reloj()
        # Una cuenta inexistente cuesta lo mismo que una real: el tiempo no delata su existencia.
        correcta = comprobar_hash(clave, fila["clave"] if fila else self._hash_ficticio)
        if fila is None:
            self.registrar(usuario, "-", "Inicio de sesión", "Cuenta inexistente", "Rechazado")
            return None
        if not fila["activo"] or fila["bloqueado_hasta"] > ahora:
            self.registrar(usuario, fila["perfil"], "Inicio de sesión", "Cuenta inhabilitada o bloqueada",
                           "Rechazado")
            return None
        if not correcta:
            intentos = fila["intentos"] + 1
            bloqueo = ahora + BLOQUEO_S if intentos >= INTENTOS_MAXIMOS else 0
            self.db.execute("UPDATE usuarios SET intentos = ?, bloqueado_hasta = ? WHERE usuario = ?",
                            (0 if bloqueo else intentos, bloqueo, usuario))
            self.db.commit()
            self.registrar(usuario, fila["perfil"], "Inicio de sesión",
                           "Bloqueo temporal" if bloqueo else "Contraseña incorrecta", "Rechazado")
            return None
        self.db.execute("UPDATE usuarios SET intentos = 0, bloqueado_hasta = 0 WHERE usuario = ?",
                        (usuario,))
        self.db.commit()
        self.registrar(usuario, fila["perfil"], "Inicio de sesión", "-", "Aceptado")
        return Sesion(usuario, fila["nombre"], fila["perfil"], ahora, bool(fila["clave_por_defecto"]))

    def sesion_valida(self, sesion):
        if sesion is None or sesion.cerrada:
            return False
        fila = self._fila(sesion.usuario)
        return bool(fila and fila["activo"] and fila["perfil"] == sesion.perfil
                    and self.reloj() - sesion.ultima_actividad < INACTIVIDAD_S)

    def actividad(self, sesion):
        if sesion is not None:
            sesion.ultima_actividad = self.reloj()

    def listar(self):
        return self.db.execute("SELECT usuario, nombre, perfil, activo, clave_por_defecto "
                               "FROM usuarios ORDER BY usuario").fetchall()

    def hay_claves_por_defecto(self):
        return bool(self.db.execute("SELECT 1 FROM usuarios WHERE clave_por_defecto = 1 AND activo = 1"
                                    " LIMIT 1").fetchone())

    def _administradores_activos(self):
        return self.db.execute("SELECT COUNT(*) FROM usuarios WHERE perfil = ? AND activo = 1",
                               (ADMINISTRADOR,)).fetchone()[0]

    def _protege_ultimo_admin(self, fila):
        if fila["perfil"] == ADMINISTRADOR and fila["activo"] and self._administradores_activos() <= 1:
            raise ErrorCuenta("No se puede dejar la celda sin una cuenta administradora activa.")

    def _exigir(self, usuario):
        fila = self._fila(usuario)
        if fila is None:
            raise ErrorCuenta("La cuenta no existe.")
        return fila

    @staticmethod
    def _validar_clave(clave):
        if len(clave) < CLAVE_MINIMA:
            raise ErrorCuenta(f"La contraseña debe tener al menos {CLAVE_MINIMA} caracteres.")

    def crear(self, usuario, nombre, perfil, clave):
        if not usuario or self._fila(usuario):
            raise ErrorCuenta("El identificador está vacío o ya existe.")
        if perfil not in PERFILES:
            raise ErrorCuenta("Perfil desconocido.")
        self._validar_clave(clave)
        self._insertar(usuario, nombre or usuario, perfil, clave)

    def cambiar_perfil(self, usuario, perfil):
        fila = self._exigir(usuario)
        if perfil not in PERFILES:
            raise ErrorCuenta("Perfil desconocido.")
        if perfil != ADMINISTRADOR:
            self._protege_ultimo_admin(fila)
        self.db.execute("UPDATE usuarios SET perfil = ? WHERE usuario = ?", (perfil, usuario))
        self.db.commit()

    def habilitar(self, usuario, activo):
        fila = self._exigir(usuario)
        if not activo:
            self._protege_ultimo_admin(fila)
        self.db.execute("UPDATE usuarios SET activo = ?, intentos = 0, bloqueado_hasta = 0 "
                        "WHERE usuario = ?", (int(activo), usuario))
        self.db.commit()

    def fijar_clave(self, usuario, clave):
        self._exigir(usuario)
        self._validar_clave(clave)
        self.db.execute("UPDATE usuarios SET clave = ?, clave_por_defecto = 0, intentos = 0, "
                        "bloqueado_hasta = 0 WHERE usuario = ?", (generar_hash(clave), usuario))
        self.db.commit()

    def cambiar_clave_propia(self, sesion, actual, nueva):
        if not comprobar_hash(actual, self._exigir(sesion.usuario)["clave"]):
            raise ErrorCuenta("La contraseña actual no es correcta.")
        self.fijar_clave(sesion.usuario, nueva)
        sesion.clave_por_defecto = False

# --- procesador.py ---

SIN_SESION = "sin sesión"

SIN_SESION_PERMITIDAS = (Op.PARADA, Op.EMERGENCIA)

@dataclass
class Resultado:
    aceptada: bool
    mensaje: str

def operativo(estado):
    return bool(estado.get("conectado") and estado.get("estacion_ok") and estado.get("coordinador"))

class Procesador:
    def __init__(self, cuentas, enviar, causas):
        self.cuentas = cuentas
        self.enviar = enviar
        self.causas = causas
        self.estado = {}
        self.pendientes = {}
        self.acks = {}

    def _registrar(self, sesion, op, detalle, resultado):
        usuario, perfil = (sesion.usuario, sesion.perfil) if sesion else (SIN_SESION, "-")
        self.cuentas.registrar(usuario, perfil, op.value, detalle, resultado)

    def _rechazar(self, sesion, op, detalle, motivo):
        self._registrar(sesion, op, detalle, "Rechazado: " + motivo)
        return Resultado(False, motivo)

    def _autorizar(self, sesion, op, detalle):
        if sesion is None and op not in SIN_SESION_PERMITIDAS:
            return self._rechazar(sesion, op, detalle, "Hace falta iniciar sesión.")
        if sesion is not None:
            if not self.cuentas.sesion_valida(sesion):
                return self._rechazar(sesion, op, detalle, "La sesión ya no es válida.")
            if not permitido(sesion.perfil, op):
                return self._rechazar(sesion, op, detalle, "El perfil no tiene este permiso.")
        return None

    def solicitar(self, sesion, op, modo=None, tipo="", senal=None, valor=None):
        detalle = self._detalle(op, modo, tipo, senal, valor)
        rechazo = self._autorizar(sesion, op, detalle)
        if rechazo:
            return rechazo
        if op in (Op.EMERGENCIA, Op.RESGUARDO, Op.REARME, Op.OBJETIVO):
            return self._seguridad(sesion, op, detalle, senal, valor)
        if op is Op.ENTRADA_SIMULADA:
            if senal not in ENTRADAS_SIMULADAS or valor not in (0, 1):
                return self._rechazar(sesion, op, detalle, "Entrada no admitida.")
            if not (self.estado.get("conectado") and self.estado.get("estacion_ok")):
                return self._rechazar(sesion, op, detalle, "Sin conexión con la estación.")
            self.enviar(("entrada", senal, valor))
            self._registrar(sesion, op, detalle, "Escrita")
            return Resultado(True, "Entrada actualizada.")
        if not operativo(self.estado):
            return self._rechazar(sesion, op, detalle, "Sin conexión con el coordinador.")
        if op is Op.ARRANQUE:
            orden, clave = ("id", "ARRANQUE_ID"), "ARRANQUE_ACK"
        elif op is Op.PARADA:
            orden, clave = ("id", "PARADA_ID"), "PARADA_ACK"
        elif op is Op.RECUPERAR:
            orden, clave = ("id", "RECUPERAR_ID"), "RECUPERAR_ACK"
        elif op is Op.REINICIAR:
            orden, clave = ("id", "REINICIAR_ID"), "REINICIAR_ACK"
        elif op is Op.PREPARAR_MODO:
            if modo not in MODOS or tipo not in TIPOS_INTERVENCION:
                return self._rechazar(sesion, op, detalle, "Selección no admitida.")
            orden, clave = ("modo", modo, False), "MODO_ACK"
        else:
            orden, clave = ("modo", 0, True), "MODO_ACK"
        self.enviar(orden)
        self.pendientes[clave] = (sesion, op, detalle)
        self._registrar(sesion, op, detalle, "Enviada")
        return Resultado(True, "Solicitud enviada; se espera la confirmación del coordinador.")

    def _seguridad(self, sesion, op, detalle, senal, valor):
        """No exige coordinador: justamente después de una parada está detenido."""
        if not (self.estado.get("conectado") and self.estado.get("estacion_ok")):
            return self._rechazar(sesion, op, detalle, "Sin conexión con la estación.")
        s = self.estado.get("senales", {})
        if op is Op.EMERGENCIA:
            if valor not in (0, 1):
                return self._rechazar(sesion, op, detalle, "Entrada no admitida.")
            self.enviar(("entrada", "EMERGENCIA_SIM", valor))
            if valor:
                self.enviar(("paro", 1))
        elif op is Op.RESGUARDO:
            if senal not in RESGUARDOS or valor not in (0, 1):
                return self._rechazar(sesion, op, detalle, "Entrada no admitida.")
            self.enviar(("entrada", senal, valor))
            # Con un modo confirmado el acceso está previsto; con equipos en marcha, detiene.
            if valor and (s.get("AUTO_ACTIVO") == 1 or s.get("MODO_EN_TRANSICION") == 1
                          or s.get("ESTADO_CONTROL") == 8):
                self.enviar(("paro", RESGUARDOS[senal]))
        elif op is Op.REARME:
            causa = s.get("PARO_CAUSA") or 0
            if not causa:
                return self._rechazar(sesion, op, detalle, "No hay una parada para rearmar.")
            if causa == 1 and sesion.perfil == PRODUCCION:
                return self._rechazar(sesion, op, detalle, "Después de una emergencia rearma mantenimiento.")
            if s.get("EMERGENCIA_SIM") == 1 or any(s.get(n) == 1 for n in RESGUARDOS):
                return self._rechazar(sesion, op, detalle, "La causa de la parada sigue presente.")
            self.enviar(("entrada", "PARO_CAUSA", 0))
        else:
            if not isinstance(valor, int) or not 0 <= valor <= OBJETIVO_MAXIMO:
                return self._rechazar(sesion, op, detalle, "Cantidad no admitida.")
            self.enviar(("entrada", "OBJETIVO_PIEZAS", valor))
        self._registrar(sesion, op, detalle, "Hecho")
        return Resultado(True, "Hecho.")

    @staticmethod
    def _detalle(op, modo, tipo, senal, valor):
        if op is Op.PREPARAR_MODO:
            return f"{tipo}: {MODOS.get(modo, modo)}"
        if op in (Op.ENTRADA_SIMULADA, Op.RESGUARDO):
            return f"{senal} = {valor}"
        if op in (Op.EMERGENCIA, Op.OBJETIVO):
            return str(valor)
        return "-"

    def actualizar(self, estado):
        """Registra la confirmación nativa, separada de la hora de la solicitud."""
        anterior, self.estado = self.estado, estado
        senales = estado.get("senales", {})
        if not operativo(estado):
            # Una orden sin confirmar no se retoma al reconectar.
            self.pendientes.clear()
            self.acks.clear()
            return
        for clave in list(self.pendientes):
            valor = senales.get(clave)
            if clave not in self.acks:
                self.acks[clave] = (anterior.get("senales", {}).get(clave, valor), False)
            base, visto = self.acks[clave]
            if visto:
                sesion, op, detalle = self.pendientes.pop(clave)
                del self.acks[clave]
                self._registrar(sesion, op, detalle, self._resultado(clave, senales))
            elif valor != base:
                self.acks[clave] = (base, True)

    def _resultado(self, clave, s):
        if clave in ("ARRANQUE_ACK", "RECUPERAR_ACK", "REINICIAR_ACK"):
            causa = int(s.get("CAUSA_RECHAZO") or 0)
            return "Confirmada" if causa == 0 else "Rechazada: " + self.causas.get(causa, str(causa))
        if clave == "MODO_ACK":
            resultado = int(s.get("MODO_RESULTADO") or 0)
            if resultado == 1:
                return "Confirmada"
            if resultado == 3:
                return "Producción detenida: reenviar la solicitud"
            causa = int(s.get("MODO_CAUSA") or 0)
            return "Rechazada: " + self.causas.get(causa, str(causa))
        return "Confirmada"

    def cerrar_sesion(self, sesion, motivo):
        """Cerrar sesión no abre la pinza ni reinicia el lote: solo pide la parada normal."""
        if sesion is None or sesion.cerrada:
            return
        sesion.cerrada = True
        detalle = motivo
        if operativo(self.estado) and self.estado.get("senales", {}).get("AUTO_ACTIVO") == 1:
            self.enviar(("id", "PARADA_ID"))
            detalle += "; parada normal solicitada"
        self.cuentas.registrar(sesion.usuario, sesion.perfil, "Cierre de sesión", detalle, "Hecho")

    def administrar(self, sesion, accion, usuario, *argumentos):
        detalle = f"{accion} {usuario}"
        rechazo = self._autorizar(sesion, Op.ADMINISTRAR, detalle)
        if rechazo:
            return rechazo
        if usuario == sesion.usuario and accion in ("cambiar_perfil", "habilitar"):
            return self._rechazar(sesion, Op.ADMINISTRAR, detalle,
                                  "Una cuenta no puede cambiar sus propios privilegios.")
        if accion not in ("crear", "cambiar_perfil", "habilitar", "fijar_clave"):
            return self._rechazar(sesion, Op.ADMINISTRAR, detalle, "Acción desconocida.")
        try:
            getattr(self.cuentas, accion)(usuario, *argumentos)
        except ErrorCuenta as error:
            return self._rechazar(sesion, Op.ADMINISTRAR, detalle, str(error))
        self._registrar(sesion, Op.ADMINISTRAR, detalle, "Hecho")
        return Resultado(True, "Cuenta actualizada.")

# --- sensores_modos.py ---

class SensoresModos:
    def __init__(self, rdk):
        self.r = rdk
        self.irb = rdk.Item("ABB IRB 1200-7/0.7", ITEM_TYPE_ROBOT)
        self.crb = rdk.Item("ABB CRB 1300-10/1.15", ITEM_TYPE_ROBOT)
        self.cinta = rdk.Item("Cinta_Pasante", ITEM_TYPE_ROBOT)
        self.tcp = rdk.Item("TCP_Pinza", ITEM_TYPE_TOOL)
        self.antorcha = rdk.Item("Antorcha_TIG", ITEM_TYPE_TOOL)
        self.targets = {n: rdk.Item(n, ITEM_TYPE_TARGET) for n in
                        ("Man_Reposo", "Sold_Reposo", "Man_Mantenimiento", "Sold_Mantenimiento",
                         "Serv_Cambio_Tungsteno")}
        self.previa = None
        self.escritos = {}
        self.estable_desde = time.monotonic()

    @staticmethod
    def cerca(q, t):
        return len(q) == len(t) and max(abs(a-b) for a,b in zip(q,t)) <= .5

    def actualizar(self):
        q = self.cinta.Joints().list()[0]
        ahora = time.monotonic()
        if self.previa is None or abs(q-self.previa) > .1:
            self.estable_desde = ahora
        self.previa = q
        # Pose real del TCP: base absoluta * cinemática directa * herramienta.
        pose = self.crb.PoseAbs() * self.crb.SolveFK(self.crb.Joints()) * self.antorcha.PoseTool()
        error = self.targets["Serv_Cambio_Tungsteno"].PoseAbs().inv() * pose
        distancia = math.sqrt(sum(v*v for v in error.Pos()))
        coseno = max(-1, min(1, (error[0,0]+error[1,1]+error[2,2]-1)/2))
        angulo = math.degrees(math.acos(coseno))
        sujeta = False
        for k in range(1,5):
            padre = self.r.Item("Estator_"+str(k)).Parent()
            while padre.Valid():
                if padre == self.tcp:
                    sujeta = True
                    break
                padre = padre.Parent()
        datos = {
            "IRB_EN_REPOSO": self.cerca(self.irb.Joints().list(), self.targets["Man_Reposo"].Joints().list()),
            "CRB_EN_REPOSO": self.cerca(self.crb.Joints().list(), self.targets["Sold_Reposo"].Joints().list()),
            "IRB_EN_MANT": self.cerca(self.irb.Joints().list(), self.targets["Man_Mantenimiento"].Joints().list()),
            "CRB_EN_MANT": self.cerca(self.crb.Joints().list(), self.targets["Sold_Mantenimiento"].Joints().list()),
            "CRB_EN_SERVICIO": distancia <= 1 and angulo <= 1,
            "CINTA_DETENIDA": ahora-self.estable_desde >= .2,
            "PIEZA_SUJETA_SENSOR": sujeta,
            "SENSORES_VALIDOS": True,
        }
        # Cada llamada a la API frena la simulación: solo se escribe lo que cambió.
        for n,v in datos.items():
            if self.escritos.get(n) != v:
                self.r.setParam(n, int(v))
                self.escritos[n] = v
        return datos

# --- enlace.py ---

ESTACION = "Celda_Soldadura_Estator_Grupo4_v05"

COORDINADOR = "Coordinador_Panel"

PERIODO_S = 0.2

REINTENTO_S = 1.0

PUERTOS = ((int(os.environ["ROBODK_API_PORT"]),) if os.environ.get("ROBODK_API_PORT")
           else (20500, 20501))

SENALES = (
    "AUTO_ACTIVO", "ESTADO_CONTROL", "CAUSA_RECHAZO", "PROXIMA_PIEZA", "PIEZA_ACTIVA",
    "PIEZAS_COMPLETADAS", "LOTES_COMPLETADOS", "ARRANQUE_ACK", "PARADA_ACK", "PARADA_ID",
    "ARCO_TIG", "MODO_ACK", "MODO_CONFIRMADO", "MODO_EN_TRANSICION", "MODO_RESULTADO",
    "MODO_CAUSA", "PERMISO_OPERACION", "IRB_DISPONIBLE", "CRB_DISPONIBLE", "CINTA_DISPONIBLE",
    "SENSORES_VALIDOS", "IRB_EN_REPOSO", "CRB_EN_REPOSO", "IRB_EN_MANT", "CRB_EN_MANT",
    "CRB_EN_SERVICIO", "CINTA_DETENIDA", "PIEZA_SUJETA_SENSOR", "PARO_CAUSA", "RECUP_PENDIENTE",
    "RECUPERAR_ACK", "REINICIAR_ACK", "EMERGENCIA_SIM", "CORTINA_ENTRADA_SIM", "CORTINA_SALIDA_SIM",
    "PUERTA_ABIERTA_SIM", "OBJETIVO_PIEZAS", "PIEZAS_BUENAS", "PIEZAS_RETRABAJO", "PEDIDOS_TERMINADOS",
    "FASE_PIEZA",
)

class RobolinkSinArranque(Robolink):
    """Robolink lanza RoboDK si no halla servidor; el panel nunca debe abrirlo por su cuenta."""

    def Connect(self):
        self.PORT = self.PORT_START
        self.NewLink()
        return 1

def puerto_abierto(puerto):
    with socket.socket() as s:
        s.settimeout(0.3)
        return s.connect_ex(("127.0.0.1", puerto)) == 0

def numero(valor):
    try:
        return float(valor)
    except (TypeError, ValueError):
        return None

class Enlace(QThread):
    estado = Signal(dict)

    def __init__(self, puertos=PUERTOS, parent=None):
        super().__init__(parent)
        self.puertos = puertos
        self.ordenes = queue.Queue()
        self.activo = True
        self.rdk = None
        self.puerto = None
        self.sensores = None
        self.estacion = None
        self.principal = None

    def enviar(self, orden):
        self.ordenes.put(orden)

    def detener(self):
        self.activo = False
        self.wait(3000)

    def _descartar_ordenes(self):
        while not self.ordenes.empty():
            self.ordenes.get_nowait()

    def _desconectar(self):
        self.rdk = self.sensores = self.estacion = self.principal = None
        self.puerto = None
        self._descartar_ordenes()

    def _conectar(self):
        for puerto in self.puertos:
            if puerto_abierto(puerto):
                self.rdk = RobolinkSinArranque(port=puerto)
                self.puerto = puerto
                return True
        return False

    def _preparar_estacion(self):
        """Devuelve True si la estación activa es la v05; rehace los ítems si fue reabierta."""
        activa = self.rdk.ActiveStation()
        if activa.Name() != ESTACION:
            self.sensores = self.estacion = self.principal = None
            self._descartar_ordenes()
            return False
        if self.estacion != activa or self.sensores is None:
            self.estacion = activa
            self.sensores = SensoresModos(self.rdk)
            self.principal = self.rdk.Item(COORDINADOR, ITEM_TYPE_PROGRAM)
        return True

    def _parar(self, causa):
        """Representa la función de seguridad: detiene sin mover nada.

        Primero el coordinador, que con una llamada frena también a sus subprogramas.
        """
        r = self.rdk
        if self.principal is not None:
            self.principal.Stop()
        for programa in r.ItemList(ITEM_TYPE_PROGRAM):
            if programa.Busy():
                programa.Stop()
        for equipo in r.ItemList(ITEM_TYPE_ROBOT):
            equipo.Stop()
        r.setParam("ARCO_TIG", 0)
        # La emergencia prevalece sobre una parada de protección que ya estuviera activa.
        if causa == 1 or not numero(r.getParam("PARO_CAUSA")):
            r.setParam("PARO_CAUSA", causa)

    def _escribir(self, orden):
        r = self.rdk
        if orden[0] == "paro":
            self._parar(orden[1])
        elif orden[0] == "id":
            senal = orden[1]
            r.setParam(senal, int(numero(r.getParam(senal)) or 0) + 1)
        elif orden[0] == "modo":
            _, modo, restitucion = orden
            if restitucion:
                r.setParam("CONF_RESTITUCION", 1)
            r.setParam("MODO_SOLICITADO", modo)
            r.setParam("MODO_ID", int(numero(r.getParam("MODO_ID")) or 0) + 1)
        elif orden[0] == "entrada":
            r.setParam(orden[1], orden[2])

    def _ciclo(self):
        if not self._preparar_estacion():
            return {"conectado": True, "estacion_ok": False, "coordinador": False,
                    "puerto": self.puerto, "senales": {}}
        self.sensores.actualizar()
        while not self.ordenes.empty():
            self._escribir(self.ordenes.get_nowait())
        valores = dict(self.rdk.getParams())
        return {"conectado": True, "estacion_ok": True, "puerto": self.puerto,
                "coordinador": bool(self.principal.Busy()),
                "senales": {n: numero(valores.get(n)) for n in SENALES}}

    def _esperar_orden(self):
        """Una orden despierta el ciclo al instante: la emergencia no espera al período."""
        limite = time.monotonic() + PERIODO_S
        while time.monotonic() < limite and self.ordenes.empty():
            time.sleep(.005)

    def run(self):
        while self.activo:
            try:
                if self.rdk is None and not self._conectar():
                    self.estado.emit({"conectado": False, "senales": {}})
                    time.sleep(REINTENTO_S)
                    continue
                self.estado.emit(self._ciclo())
                self._esperar_orden()
            except Exception:
                # Caída de RoboDK o estación cerrada a mitad de una consulta.
                self._desconectar()
                self.estado.emit({"conectado": False, "senales": {}})
                time.sleep(REINTENTO_S)
        try:
            if self.sensores is not None:
                # Cerrar el panel en producción encola una parada que debe salir antes de terminar.
                while not self.ordenes.empty():
                    self._escribir(self.ordenes.get_nowait())
                self.rdk.setParam("SENSORES_VALIDOS", 0)
        except Exception:
            pass

# --- sinoptico.py ---

X_MIN, X_MAX, Y_MIN, Y_MAX = -2150.0, 2200.0, -1250.0, 2150.0

CERRAMIENTO = (-1300.0, 850.0, -960.0, 1850.0)

BANDA = (-2000.0, 2100.0, -860.0, -260.0)

PUERTA_Y = (1000.0, 1700.0)

CORTINA_Y = (-960.0, -120.0)

IRB = (0.0, 0.0)

CRB = (0.0, 1150.0)

PULSADORES = ((930.0, 920.0), (-1420.0, -1060.0), (970.0, -1060.0), (1150.0, 250.0))

FONDO = QColor("#f8f9fa")

LINEA = QColor("#3a4651")

NORMAL = QColor("#1d6b45")

ALERTA = QColor("#b3261e")

BANDA_C = QColor("#55606a")

ROBOT = QColor("#dfe5ea")

class Sinoptico(QWidget):
    accionado = Signal(str)

    def __init__(self, parent=None):
        super().__init__(parent)
        self.senales = {}
        self.zonas = {}
        self.setMinimumSize(420, 340)
        self.setSizePolicy(QSizePolicy.Expanding, QSizePolicy.Expanding)
        self.setCursor(Qt.PointingHandCursor)

    def actualizar(self, senales):
        self.senales = senales
        self.update()

    def _escala(self):
        return min(self.width() / (X_MAX - X_MIN), self.height() / (Y_MAX - Y_MIN))

    def _punto(self, x, y):
        e = self._escala()
        margen_x = (self.width() - (X_MAX - X_MIN) * e) / 2
        margen_y = (self.height() - (Y_MAX - Y_MIN) * e) / 2
        return QPointF(margen_x + (x - X_MIN) * e, margen_y + (Y_MAX - y) * e)

    def _rect(self, x0, x1, y0, y1):
        return QRectF(self._punto(x0, y1), self._punto(x1, y0))

    def _activa(self, senal):
        return self.senales.get(senal) == 1

    def _texto(self, p, x, y, texto, color=LINEA, negrita=False):
        fuente = QFont("Segoe UI", 8)
        fuente.setBold(negrita)
        p.setFont(fuente)
        p.setPen(color)
        punto = self._punto(x, y)
        p.drawText(QRectF(punto.x() - 90, punto.y() - 10, 180, 20), Qt.AlignCenter, texto)

    def _cortina(self, p, nombre, senal, x, etiqueta, texto_x):
        cortada = self._activa(senal)
        color = ALERTA if cortada else NORMAL
        p.setPen(QPen(color, 4, Qt.DashLine))
        p.drawLine(self._punto(x, CORTINA_Y[0]), self._punto(x, CORTINA_Y[1]))
        self._texto(p, texto_x, CORTINA_Y[1] + 120, f"{etiqueta}: {'cortada' if cortada else 'libre'}", color, True)
        self.zonas[nombre] = self._rect(min(x, texto_x) - 500, max(x, texto_x) + 500 if texto_x > x else x + 170,
                                        CORTINA_Y[0], CORTINA_Y[1] + 240)

    def _robot(self, p, posicion, nombre, reposo, mantenimiento):
        centro = self._punto(*posicion)
        radio = 330 * self._escala()
        p.setPen(QPen(LINEA, 1.5))
        p.setBrush(QBrush(ROBOT))
        p.drawEllipse(centro, radio, radio)
        estado = "reposo" if self._activa(reposo) else "mantenimiento" if self._activa(mantenimiento) else "en ciclo"
        self._texto(p, posicion[0], posicion[1] + 50, nombre, LINEA, True)
        self._texto(p, posicion[0], posicion[1] - 90, estado)

    def paintEvent(self, _):
        p = QPainter(self)
        p.setRenderHint(QPainter.Antialiasing)
        p.fillRect(self.rect(), FONDO)
        self.zonas = {}
        x0, x1, y0, y1 = CERRAMIENTO
        p.setPen(QPen(LINEA, 2))
        p.setBrush(Qt.NoBrush)
        p.drawRect(self._rect(x0, x1, y0, y1))
        p.setPen(Qt.NoPen)
        p.setBrush(QBrush(BANDA_C))
        p.drawRect(self._rect(*BANDA))
        self._texto(p, -500, -560, "Cinta", QColor("#ffffff"), True)

        self._robot(p, IRB, "IRB 1200", "IRB_EN_REPOSO", "IRB_EN_MANT")
        self._robot(p, CRB, "CRB 1300", "CRB_EN_REPOSO", "CRB_EN_MANT")
        if self._activa("ARCO_TIG"):
            self._texto(p, 500, 650, "ARCO ENCENDIDO", ALERTA, True)

        self._cortina(p, "cortina_entrada", "CORTINA_ENTRADA_SIM", x0, "Cortina entrada", x0 - 620)
        self._cortina(p, "cortina_salida", "CORTINA_SALIDA_SIM", x1, "Cortina salida", x1 + 620)

        abierta = self._activa("PUERTA_ABIERTA_SIM")
        color = ALERTA if abierta else NORMAL
        p.setPen(QPen(color, 6))
        bisagra = self._punto(x1, PUERTA_Y[0])
        if abierta:
            p.drawLine(bisagra, self._punto(x1 + 620, PUERTA_Y[0] + 320))
        else:
            p.drawLine(bisagra, self._punto(x1, PUERTA_Y[1]))
        self._texto(p, x1 + 620, PUERTA_Y[1] + 110, f"Puerta: {'abierta' if abierta else 'cerrada'}", color, True)
        self.zonas["puerta"] = self._rect(x1 - 150, x1 + 800, PUERTA_Y[0] - 100, PUERTA_Y[1] + 200)

        pulsado = self._activa("EMERGENCIA_SIM")
        radio = 75 * self._escala() + 5
        for i, posicion in enumerate(PULSADORES):
            centro = self._punto(*posicion)
            p.setPen(QPen(QColor("#d9a400"), 3))
            p.setBrush(QBrush(ALERTA if pulsado else QColor("#d8453c")))
            p.drawEllipse(centro, radio, radio)
            self.zonas[f"emergencia_{i}"] = QRectF(centro.x() - radio - 4, centro.y() - radio - 4,
                                                   2 * radio + 8, 2 * radio + 8)
        p.end()

    def mousePressEvent(self, evento):
        # Las zonas de los pulsadores tienen prioridad: están dentro de otras.
        for nombre, zona in sorted(self.zonas.items(), key=lambda z: not z[0].startswith("emergencia")):
            if zona.contains(evento.pos()):
                self.accionado.emit("emergencia" if nombre.startswith("emergencia") else nombre)
                return

# --- ventana.py ---

ESTADOS = {0: "Inicial", 1: "Automático", 2: "Parada normal", 3: "Detenida por condición perdida",
           4: "Preparando modo", 5: "Regresando de modo", 6: "Modo confirmado",
           7: "Recuperación pendiente", 8: "Recuperando", 9: "Pedido terminado"}

FASES = {1: "avance", 2: "toma", 3: "presentación", 4: "soldadura", 5: "giro", 6: "soldadura", 7: "depósito",
         8: "regreso"}

RESULTADOS_MODO = {1: "Aceptada", 2: "Rechazada", 3: "Producción detenida: reenviar la solicitud"}

SENSORES = (("IRB_EN_REPOSO", "IRB en reposo"), ("CRB_EN_REPOSO", "CRB en reposo"),
            ("IRB_EN_MANT", "IRB en mantenimiento"), ("CRB_EN_MANT", "CRB en mantenimiento"),
            ("CRB_EN_SERVICIO", "CRB en servicio"), ("CINTA_DETENIDA", "Cinta detenida"),
            ("PIEZA_SUJETA_SENSOR", "Pieza sujeta"), ("SENSORES_VALIDOS", "Sensores en ejecución"))

ETIQUETAS_ENTRADA = {"PERMISO_OPERACION": "Permiso de operación", "IRB_DISPONIBLE": "IRB disponible",
                     "CRB_DISPONIBLE": "CRB disponible", "CINTA_DISPONIBLE": "Cinta disponible"}

AYUDA = """
<h3>Cómo usar la celda</h3>
<p><b>Ciclo completo sin panel:</b> doble clic en <code>Programa_Principal</code>. Suelda un lote de
cuatro estatores y termina.</p>
<p><b>Con el panel:</b></p>
<ol>
<li>Doble clic en <code>Coordinador_Panel</code>: queda esperando órdenes y nada se mueve.</li>
<li>Doble clic en <code>Panel_Operador</code>, si no está abierto.</li>
<li>Entrar como mantenimiento y marcar las cuatro entradas de simulación.</li>
<li>Cerrar sesión, entrar como producción y pulsar Arranque.</li>
</ol>
<p>No mezclar: para pasar de un programa a otro, reabrir la estación sin guardar.</p>
<h3>Paradas</h3>
<p><b>Emergencia:</b> botón rojo de la banda o pulsadores de la pestaña Proceso. <b>Cortinas y puerta:</b>
clic en la imagen del proceso; detienen solo si hay equipos en marcha.</p>
<p>Después de una parada: eliminar la causa, pulsar Rearme, doble clic en <code>Coordinador_Panel</code> y,
si la pieza quedó a medias, Recuperar con mantenimiento. Una pieza cortada al soldar se termina y se
deja corrida en la cinta, como retrabajo. Rearmar no arranca nada.</p>
<h3>Cantidad a fabricar</h3>
<p>En Producción, fijar el objetivo de piezas buenas; 0 es sin límite. El retrabajo no cuenta. Al llegar,
la celda repone las piezas, pone los contadores en cero y queda lista.</p>
<h3>Cuentas de puesta en marcha</h3>
{cuentas}
<h3>Perfiles</h3>
<ul>
<li><b>Producción:</b> arranque, parada, objetivo y rearme de cortinas y puerta.</li>
<li><b>Mantenimiento:</b> modos, entradas de simulación, rearme, recuperación y reinicio de lote.</li>
<li><b>Administrador:</b> cuentas y parada; no opera la celda.</li>
</ul>
<h3>Mantenimiento</h3>
<p>Elegir equipo y pulsar Preparar. Si había producción, se detiene al terminar la pieza: pulsar
Preparar otra vez. Al terminar, Confirmar restitución y regresar; la celda no arranca sola.</p>
<h3>Límites</h3>
<ul>
<li>Parada normal termina la pieza en curso: no es una parada de emergencia.</li>
<li>La emergencia del panel representa la función: la real es un circuito de seguridad.</li>
<li>Las entradas de simulación no son protecciones.</li>
<li>El panel solo envía solicitudes: los movimientos son programas nativos de RoboDK.</li>
<li>Al cerrar RoboDK, no guardar: se conservaría el estado de la simulación.</li>
</ul>
"""

ESTILO = """
QMainWindow, QWidget#fondo { background: #eef0f2; }
QWidget { color: #1c2329; font-family: "Segoe UI"; font-size: 14px; }
QFrame#banda { background: #1f2d3a; }
QFrame#banda QLabel { color: #ffffff; }
QLabel#titulo { font-size: 17px; font-weight: 600; }
QFrame#tarjeta, QGroupBox { background: #ffffff; border: 1px solid #cfd5da; border-radius: 6px; }
QGroupBox { margin-top: 14px; padding-top: 12px; font-weight: 600; }
QGroupBox::title { subcontrol-origin: margin; left: 10px; padding: 0 4px; }
QLabel#rotulo { color: #56626c; font-size: 12px; }
QLabel#valor { font-size: 15px; font-weight: 600; }
QLabel#aviso { background: #fff3cd; border: 1px solid #d9b64a; border-radius: 4px; padding: 6px 10px; }
QLabel#mensaje { color: #1c2329; padding: 2px; }
QPushButton { background: #ffffff; border: 1px solid #8b98a3; border-radius: 4px; padding: 7px 14px; }
QPushButton:hover { background: #e4e9ed; }
QPushButton:disabled { color: #8f99a1; border-color: #cfd5da; background: #f2f4f5; }
QPushButton#primario, QPushButton#crear_cuenta { background: #1d6b45; border-color: #1d6b45; color: #ffffff; font-weight: 600; }
QPushButton#primario:disabled { background: #c9d6cf; border-color: #c9d6cf; color: #ffffff; }
QPushButton#parada { background: #b3261e; border-color: #b3261e; color: #ffffff; font-weight: 600; }
QPushButton#parada:disabled { background: #dcbcba; border-color: #dcbcba; color: #ffffff; }
QPushButton#emergencia { background: #ffcc00; border: 3px solid #b3261e; color: #b3261e; font-weight: 700; }
QPushButton#emergencia:disabled { background: #efe6bd; border-color: #d9c9a0; color: #a89b6d; }
QTabWidget::pane { border: 1px solid #cfd5da; background: #f8f9fa; }
QTabBar::tab { padding: 8px 18px; background: #dfe3e7; border: 1px solid #cfd5da; }
QTabBar::tab:selected { background: #f8f9fa; color: #1d6b45; }
QTableWidget { background: #ffffff; gridline-color: #e1e5e8; }
QLineEdit, QComboBox, QSpinBox { background: #ffffff; border: 1px solid #8b98a3; border-radius: 4px; padding: 5px; }
"""

def rotulo(texto):
    etiqueta = QLabel(texto)
    etiqueta.setObjectName("rotulo")
    etiqueta.setWordWrap(True)
    return etiqueta

def tarjeta(titulo):
    marco = QFrame()
    marco.setObjectName("tarjeta")
    capa = QVBoxLayout(marco)
    capa.setContentsMargins(12, 8, 12, 8)
    capa.addWidget(rotulo(titulo))
    valor = QLabel("—")
    valor.setObjectName("valor")
    valor.setWordWrap(True)
    valor.setMinimumHeight(48)
    valor.setAlignment(Qt.AlignLeft | Qt.AlignTop)
    capa.addWidget(valor)
    return marco, valor

def tabla(columnas):
    t = QTableWidget(0, len(columnas))
    t.setHorizontalHeaderLabels(columnas)
    t.verticalHeader().hide()
    t.setEditTriggers(QAbstractItemView.NoEditTriggers)
    t.setSelectionBehavior(QAbstractItemView.SelectRows)
    t.horizontalHeader().setSectionResizeMode(QHeaderView.Stretch)
    return t

def llenar(t, filas):
    t.setRowCount(len(filas))
    for i, fila in enumerate(filas):
        for j, valor in enumerate(fila):
            t.setItem(i, j, QTableWidgetItem(str(valor)))

def condiciones_arranque(s):
    """Solo para mostrar; quien decide es el coordinador nativo."""
    igual = lambda n, v: s.get(n) == v
    return (("Permiso de operación", igual("PERMISO_OPERACION", 1)),
            ("Sensores en ejecución", igual("SENSORES_VALIDOS", 1)),
            ("Sin modo activo", igual("MODO_CONFIRMADO", 0) and igual("MODO_EN_TRANSICION", 0)),
            ("Robots en reposo", igual("IRB_EN_REPOSO", 1) and igual("CRB_EN_REPOSO", 1)),
            ("Sin pieza sujeta", igual("PIEZA_SUJETA_SENSOR", 0)),
            ("Sin parada activa", not s.get("PARO_CAUSA")),
            ("Resguardos cerrados", not any(igual(n, 1) for n in RESGUARDOS)),
            ("Sin recuperación pendiente", igual("RECUP_PENDIENTE", 0)),
            ("Cinta detenida", igual("CINTA_DETENIDA", 1)),
            ("Equipos disponibles", igual("IRB_DISPONIBLE", 1) and igual("CRB_DISPONIBLE", 1)
             and igual("CINTA_DISPONIBLE", 1)))

class Ventana(QMainWindow):
    def __init__(self, cuentas, procesador, causas, version="v05"):
        super().__init__()
        self.cuentas = cuentas
        self.procesador = procesador
        self.causas = causas
        self.sesion = None
        self.estado = {}
        self.setWindowTitle(f"Panel de operador · Celda de soldadura TIG {version}")
        self.resize(1040, 720)
        self.setStyleSheet(ESTILO)
        fondo = QWidget()
        fondo.setObjectName("fondo")
        self.setCentralWidget(fondo)
        capa = QVBoxLayout(fondo)
        capa.setContentsMargins(0, 0, 0, 0)
        capa.addWidget(self._banda())
        cuerpo = QVBoxLayout()
        cuerpo.setContentsMargins(14, 10, 14, 12)
        cuerpo.addLayout(self._resumen())
        self.aviso = QLabel()
        self.aviso.setObjectName("aviso")
        self.aviso.setWordWrap(True)
        self.aviso.hide()
        cuerpo.addWidget(self.aviso)
        self.paginas = QStackedWidget()
        self.paginas.addWidget(self._pagina_login())
        self.pestanas = QTabWidget()
        self.paginas.addWidget(self.pestanas)
        cuerpo.addWidget(self.paginas, 1)
        capa.addLayout(cuerpo, 1)
        self._construir_pestanas()
        self.reloj = QTimer(self)
        self.reloj.timeout.connect(self._vigilar_sesion)
        self.reloj.start(1000)
        self._refrescar_sesion()

    # Construcción

    def _banda(self):
        banda = QFrame()
        banda.setObjectName("banda")
        capa = QHBoxLayout(banda)
        capa.setContentsMargins(14, 8, 14, 8)
        titulo = QLabel("Panel")
        titulo.setObjectName("titulo")
        capa.addWidget(titulo)
        capa.addStretch(1)
        self.et_conexion = QLabel()
        capa.addWidget(self.et_conexion)
        capa.addSpacing(18)
        self.et_usuario = QLabel()
        capa.addWidget(self.et_usuario)
        self.bt_ayuda = QPushButton("Ayuda")
        self.bt_ayuda.clicked.connect(self._ayuda)
        capa.addWidget(self.bt_ayuda)
        self.bt_clave = QPushButton("Contraseña")
        self.bt_clave.clicked.connect(self._cambiar_clave)
        capa.addWidget(self.bt_clave)
        self.bt_salir = QPushButton("Cerrar sesión")
        self.bt_salir.clicked.connect(lambda: self._cerrar_sesion("Cierre por el usuario"))
        capa.addWidget(self.bt_salir)
        self.bt_parada = QPushButton("Parada normal")
        self.bt_parada.setObjectName("parada")
        self.bt_parada.clicked.connect(lambda: self._orden(Op.PARADA))
        capa.addWidget(self.bt_parada)
        self.bt_emergencia = QPushButton("EMERGENCIA")
        self.bt_emergencia.setObjectName("emergencia")
        self.bt_emergencia.clicked.connect(self._alternar_emergencia)
        capa.addWidget(self.bt_emergencia)
        return banda

    def _resumen(self):
        fila = QHBoxLayout()
        self.valores = {}
        for clave, titulo in (("estado", "Estado de la celda"), ("modo", "Modo confirmado"),
                              ("pieza", "Pieza y lote"), ("causa", "Último rechazo")):
            marco, valor = tarjeta(titulo)
            self.valores[clave] = valor
            fila.addWidget(marco, 1)
        return fila

    def _pagina_login(self):
        pagina = QWidget()
        externa = QGridLayout(pagina)
        caja = QGroupBox("Inicio de sesión")
        caja.setMinimumWidth(360)
        formulario = QFormLayout(caja)
        self.in_usuario = QLineEdit()
        self.in_clave = QLineEdit()
        self.in_clave.setEchoMode(QLineEdit.Password)
        self.in_clave.returnPressed.connect(self._entrar)
        formulario.addRow("Usuario", self.in_usuario)
        formulario.addRow("Contraseña", self.in_clave)
        self.bt_entrar = QPushButton("Entrar")
        self.bt_entrar.setObjectName("primario")
        self.bt_entrar.clicked.connect(self._entrar)
        formulario.addRow(self.bt_entrar)
        self.et_login = QLabel()
        self.et_login.setWordWrap(True)
        formulario.addRow(self.et_login)
        externa.addWidget(caja, 0, 0, Qt.AlignCenter)
        return pagina

    def _pestana_produccion(self):
        pagina = QWidget()
        capa = QHBoxLayout(pagina)
        mandos = QGroupBox("Mandos")
        columna = QVBoxLayout(mandos)
        self.bt_arranque = QPushButton("Arranque")
        self.bt_arranque.setObjectName("primario")
        self.bt_arranque.clicked.connect(lambda: self._orden(Op.ARRANQUE))
        columna.addWidget(self.bt_arranque)
        self.et_arranque = QLabel()
        self.et_arranque.setWordWrap(True)
        columna.addWidget(self.et_arranque)
        columna.addWidget(rotulo("La parada normal termina y deposita la pieza en curso. "
                                 "No es una parada de emergencia."))
        fila = QHBoxLayout()
        fila.addWidget(QLabel("Piezas buenas a fabricar"))
        self.sp_objetivo = QSpinBox()
        self.sp_objetivo.setRange(0, OBJETIVO_MAXIMO)
        self.sp_objetivo.setSpecialValueText("Sin límite")
        fila.addWidget(self.sp_objetivo)
        self.bt_objetivo = QPushButton("Fijar")
        self.bt_objetivo.clicked.connect(lambda: self._orden(Op.OBJETIVO, self.et_arranque,
                                                             valor=self.sp_objetivo.value()))
        fila.addWidget(self.bt_objetivo)
        columna.addLayout(fila)
        columna.addWidget(rotulo("El retrabajo no cuenta. Al llegar, la celda repone las piezas y "
                                 "pone los contadores en cero."))
        columna.addStretch(1)
        capa.addWidget(mandos, 1)
        caja = QGroupBox("Condiciones de arranque")
        lista = QVBoxLayout(caja)
        self.et_condiciones = QLabel()
        self.et_condiciones.setTextFormat(Qt.PlainText)
        lista.addWidget(self.et_condiciones)
        lista.addStretch(1)
        capa.addWidget(caja, 1)
        return pagina

    def _pestana_mantenimiento(self):
        pagina = QWidget()
        capa = QHBoxLayout(pagina)
        caja = QGroupBox("Preparación")
        formulario = QFormLayout(caja)
        self.cb_modo = QComboBox()
        for modo, nombre in MODOS.items():
            self.cb_modo.addItem(nombre, modo)
        self.cb_tipo = QComboBox()
        self.cb_tipo.addItems(TIPOS_INTERVENCION)
        formulario.addRow("Equipo o tarea", self.cb_modo)
        formulario.addRow("Intervención", self.cb_tipo)
        self.bt_preparar = QPushButton("Preparar")
        self.bt_preparar.setObjectName("primario")
        self.bt_preparar.clicked.connect(self._preparar)
        formulario.addRow(self.bt_preparar)
        self.bt_regresar = QPushButton("Confirmar restitución y regresar")
        self.bt_regresar.clicked.connect(self._regresar)
        formulario.addRow(self.bt_regresar)
        self.et_modo = QLabel()
        self.et_modo.setWordWrap(True)
        formulario.addRow(self.et_modo)
        formulario.addRow(rotulo("La preparación posiciona los equipos. El aislamiento y el bloqueo "
                                 "se hacen por procedimiento, fuera del panel; esta confirmación "
                                 "no es una medición de energía cero."))
        capa.addWidget(caja, 3)
        simuladas = QGroupBox("Entradas de simulación")
        columna = QVBoxLayout(simuladas)
        columna.addWidget(rotulo("Representan señales externas de la celda. No son protecciones."))
        self.entradas = {}
        for senal in ENTRADAS_SIMULADAS:
            casilla = QCheckBox(ETIQUETAS_ENTRADA[senal])
            # PySide2 no pasa el argumento de clicked a una lambda con valores por defecto.
            casilla.clicked.connect(lambda _=False, s=senal, c=casilla: self._entrada(s, c.isChecked()))
            self.entradas[senal] = casilla
            columna.addWidget(casilla)
        columna.addStretch(1)
        capa.addWidget(simuladas, 2)
        return pagina

